(* IEC 61131-3 sources: daoli-st-library/DL_Device (part 18) *)

(* ---- FB_DL_CrystallizerVacuumCtrl.st ---- *)
(*
  Component : FB_DL_CrystallizerVacuumCtrl
  Category  : DL_Device
  Type      : FB
  Complexity: C2
  VERSION   : v1.0.0
  功能      : 结晶罐真空控制：ENUM 四态（Off/Run/Lost/Fault），真空泵按压差分级投运，按锤度算沸点升高与罐内沸点，真空丢失延时联锁停泵。
  开源溯源  : 道莅原创 clean-room 自研（无外部代码引用）｜License: MIT
  边界条件  : ① 真空度输入按罐内绝对压力定义 [kPa]：实测值升高即真空丢失，判据方向不得反接；
              ② 沸点升高按 锤度/(100-锤度) 经验式，锤度须 < 100 °Bx 且钳位 0~30 K；
              ③ 真空丢失锁存后全泵切除（防倒吸油返），唯一解除路径 = bReset 上升沿。
*)

TYPE E_DL_VacMode :
(
    eOff   := 0,    (* 停机：使能撤销 / Off, disabled *)
    eRun   := 10,   (* 运行：分级投运 / Running with staged pumps *)
    eLost  := 20,   (* 真空丢失：全泵切除锁存 / Vacuum lost, pumps cut off *)
    eFault := 90    (* 故障：锁存待复位 / Fault latched *)
);
END_TYPE

FUNCTION_BLOCK FB_DL_CrystallizerVacuumCtrl
VAR_INPUT
    bEnable     : BOOL;   (* 使能电平 [-] Enable level *)
    bReset      : BOOL;   (* 复位上升沿，清丢失与故障锁存 [-] Reset edge *)
    fVacuumKPa  : REAL;   (* 罐内绝对压力实测 [kPa] Measured absolute pressure *)
    fVacSetKPa  : REAL;   (* 目标绝对压力设定 [kPa] Absolute pressure setpoint *)
    fVacLostKPa : REAL;   (* 真空丢失判据压力 [kPa] Vacuum-lost pressure threshold *)
    fBrixPct    : REAL;   (* 糖膏锤度 [°Bx] Massecuite brix *)
    fWaterBoilC : REAL;   (* 当前真空下纯水沸点 [°C] Water boiling point at this vacuum *)
    tLostDelay  : TIME;   (* 真空丢失确认延时 [ms] Vacuum-lost confirmation delay *)
    nPumpMax    : INT;    (* 可用真空泵台数 1~3 [-] Available pump count *)
END_VAR
VAR_OUTPUT
    abPumpCmd  : ARRAY[0..2] OF BOOL;  (* 三级真空泵指令 [-] Vacuum pump commands *)
    nPumpRun   : INT;                  (* 当前投运泵台数 [-] Running pump count *)
    fBoilRiseK : REAL;                 (* 沸点升高 [K] Boiling point elevation *)
    fBoilTempC : REAL;                 (* 罐内糖膏沸点 [°C] Massecuite boiling point *)
    bVacLost   : BOOL;                 (* 真空丢失锁存标志 [-] Vacuum lost latch *)
    eMode      : E_DL_VacMode;         (* 模式出口，段尾单点映射 [-] Mode outlet *)
    bError     : BOOL;                 (* 故障锁存标志 [-] Fault latch flag *)
    uErrId     : UDINT;                (* 事件码，0 = 无事件 [-] Event code *)
END_VAR
VAR
    rtReset  : R_TRIG;   (* 复位沿实例，每拍无条件刷新 / Reset edge *)
    tonLost  : TON;      (* 真空丢失确认计时 / Vacuum lost timer *)
    _eMode   : E_DL_VacMode := E_DL_VacMode.eOff;  (* 内部模式 / Internal mode *)
    _bLost   : BOOL;     (* 真空丢失锁存位（锁存量） / Latched vacuum lost bit *)
    _bFault  : BOOL;     (* 故障锁存位（锁存量） / Latched fault bit *)
    _uFault  : UDINT;    (* 故障码锁存（锁存量） / Latched fault code *)
    _bCfgBad : BOOL;     (* 组态非法当拍量 [-] Config illegal flag *)
    _bNonFin : BOOL;     (* 输入非有限当拍量 [-] Non-finite input flag *)
    nIdx     : INT;      (* 泵组遍历下标 [-] Pump loop index *)
    fErrKPa  : REAL;     (* 压差（实测 - 设定） [kPa] Pressure error *)
    fDenBrix : REAL;     (* 锤度余量（100 - 锤度） [°Bx] Brix headroom *)
END_VAR
VAR CONSTANT
    DL_EPS      : REAL := 1.0E-9;   (* 除零判定容差 [无量纲] Divide-by-zero tolerance *)
    DL_BAND1    : REAL := 1.0;      (* 一级投运压差 [kPa] Stage 1 pressure band *)
    DL_BAND2    : REAL := 4.0;      (* 二级投运压差 [kPa] Stage 2 pressure band *)
    DL_BAND3    : REAL := 8.0;      (* 三级投运压差 [kPa] Stage 3 pressure band *)
    DL_RISE_K   : REAL := 2.6;      (* 沸点升高经验系数 [K] Elevation coefficient *)
    DL_RISE_MAX : REAL := 30.0;     (* 沸点升高上限 [K] Elevation upper clamp *)
    DL_PCT_BASE : REAL := 100.0;    (* 百分比基准 [°Bx 基准] Percent base *)
    DL_IDX_MAX  : INT := 2;         (* 泵组最高下标 [-] Highest pump index *)
END_VAR

(* —— 段 0｜沿与定时器每拍无条件刷新（禁置于 IF/CASE 内，使能挂 IN 引脚） —— *)
rtReset(CLK := bReset);
tonLost(IN := bEnable AND (fVacuumKPa >= fVacLostKPa) AND (NOT _bLost), PT := tLostDelay);

(* —— 段 1｜每拍量预清零 + 泵指令全预置（锁存量 _bLost/_bFault/_uFault 不入清单） —— *)
uErrId := 16#0000_0000;
_bCfgBad := FALSE;
_bNonFin := FALSE;
nPumpRun := 0;
FOR nIdx := 0 TO 2 DO
    IF (nIdx >= 0) AND (nIdx <= DL_IDX_MAX) THEN
        abPumpCmd[nIdx] := FALSE;            (* 泵指令预置停止 [-] / Pump preset off *)
    END_IF
END_FOR

(* —— 段 2｜非有限拦截与组态闸（覆盖压力设定/丢失判据/锤度/延时/泵数） —— *)
IF (fVacuumKPa <> fVacuumKPa) OR ((fVacuumKPa - fVacuumKPa) <> 0.0)
   OR (fBrixPct <> fBrixPct) OR ((fBrixPct - fBrixPct) <> 0.0)
   OR (fVacSetKPa <> fVacSetKPa) OR ((fVacSetKPa - fVacSetKPa) <> 0.0)
   OR (fVacLostKPa <> fVacLostKPa) OR ((fVacLostKPa - fVacLostKPa) <> 0.0)
   OR (fWaterBoilC <> fWaterBoilC) OR ((fWaterBoilC - fWaterBoilC) <> 0.0) THEN
    _bNonFin := TRUE;
END_IF
IF (fVacSetKPa <= DL_EPS) OR (fVacLostKPa <= fVacSetKPa) OR (tLostDelay = T#0S)
   OR (nPumpMax < 1) OR (nPumpMax > 3) OR (fBrixPct < 0.0) OR (fBrixPct >= DL_PCT_BASE) THEN
    _bCfgBad := TRUE;
END_IF

(* —— 段 3｜沸点升高与罐内沸点：dT = 2.6·B/(100-B)，钳位 0~30 K —— *)
fDenBrix := DL_PCT_BASE - fBrixPct;
IF fDenBrix > DL_EPS THEN
    fBoilRiseK := DL_RISE_K * fBrixPct / fDenBrix;
ELSE
    fBoilRiseK := DL_RISE_MAX;               (* 锤度近饱和：按上限处理 *)
END_IF
IF fBoilRiseK < 0.0 THEN
    fBoilRiseK := 0.0;
ELSIF fBoilRiseK > DL_RISE_MAX THEN
    fBoilRiseK := DL_RISE_MAX;
END_IF
fBoilTempC := fWaterBoilC + fBoilRiseK;

(* —— 段 4｜复位沿：一次性清丢失与故障锁存（唯一解除路径，恒可达） —— *)
IF rtReset.Q THEN
    _bLost := FALSE;
    _bFault := FALSE;
    _uFault := 16#0000_0000;
    _eMode := E_DL_VacMode.eOff;
END_IF
IF _bCfgBad AND (NOT _bFault) THEN
    _bFault := TRUE;
    _uFault := 16#0029_0001;                 (* 故障级：组态非法 / Fault code bad config *)
END_IF
IF _bNonFin AND (NOT _bFault) THEN
    _bFault := TRUE;
    _uFault := 16#0029_0002;                 (* 故障级：压力或锤度非有限 / Non-finite input *)
END_IF
IF tonLost.Q AND (NOT _bLost) THEN
    _bLost := TRUE;                          (* 真空丢失锁存：全泵切除防倒吸 *)
END_IF

(* —— 段 5｜模式机：四态全覆盖 + ELSE 兜底 —— *)
CASE _eMode OF
E_DL_VacMode.eOff:
    nPumpRun := 0;
    IF bEnable AND (NOT _bLost) AND (NOT _bFault) AND (NOT _bCfgBad) AND (NOT _bNonFin) THEN
        _eMode := E_DL_VacMode.eRun;         (* 迁入条件：使能且无任何锁存 *)
    END_IF

E_DL_VacMode.eRun:
    (* 压差分级投运：实测绝对压力高于设定越多，投运泵台数越多 *)
    fErrKPa := fVacuumKPa - fVacSetKPa;
    IF fErrKPa > DL_BAND3 THEN
        nPumpRun := 3;
    ELSIF fErrKPa > DL_BAND2 THEN
        nPumpRun := 2;
    ELSIF fErrKPa > DL_BAND1 THEN
        nPumpRun := 1;
    ELSE
        nPumpRun := 0;
    END_IF
    IF nPumpRun > nPumpMax THEN
        nPumpRun := nPumpMax;                (* 受可用台数限制 [-] / Limited by available pumps *)
    END_IF
    IF _bLost THEN
        _eMode := E_DL_VacMode.eLost;        (* 迁出条件 1：真空丢失 *)
    ELSIF _bFault THEN
        _eMode := E_DL_VacMode.eFault;       (* 迁出条件 2：故障锁存 *)
    ELSIF NOT bEnable THEN
        _eMode := E_DL_VacMode.eOff;         (* 迁出条件 3：使能撤销 *)
    END_IF

E_DL_VacMode.eLost:
    nPumpRun := 0;                           (* 丢失相：全泵切除（防倒吸油返） *)
    IF NOT _bLost THEN
        _eMode := E_DL_VacMode.eOff;         (* 迁出条件：锁存被复位沿清除 *)
    END_IF

E_DL_VacMode.eFault:
    nPumpRun := 0;                           (* 故障相：全泵切除 *)
    IF (NOT _bFault) AND (NOT _bLost) THEN
        _eMode := E_DL_VacMode.eOff;         (* 迁出条件：故障锁存被复位沿清除 *)
    END_IF

ELSE
    _bFault := TRUE;                         (* 兜底：非法模式锁存 *)
    _uFault := 16#0029_0009;
    _eMode := E_DL_VacMode.eFault;
END_CASE

(* —— 段 6｜泵指令下发：仅运行相按台数投运，其余相全切除 —— *)
IF _eMode = E_DL_VacMode.eRun THEN
    FOR nIdx := 0 TO 2 DO
        IF (nIdx >= 0) AND (nIdx <= DL_IDX_MAX) THEN
            abPumpCmd[nIdx] := nIdx < nPumpRun;   (* 前 nPumpRun 台投运 [-] / First N pumps on *)
        END_IF
    END_FOR
ELSE
    nPumpRun := 0;
END_IF

(* —— 段 7｜出口单点映射 —— *)
eMode := _eMode;
bVacLost := _bLost;
bError := _bFault;
IF _bFault AND (_uFault <> 16#0000_0000) THEN
    uErrId := _uFault;                       (* 故障码锁存回放 / Latched fault replay *)
END_IF
END_FUNCTION_BLOCK

(* ---- FB_DL_CurtainEFEMZone.st ---- *)
(*
  FB_DL_CurtainEFEMZone  —  EFEM 区内光幕分区（四路遮光判向 / 屏蔽窗管理 / 顺序故障锁存）/ EFEM zone light-curtain muting
  分类 Category : DL_Device
  码位 Code     : 16#03_2_0C
  版本 Version  : 1.0.2
  来源 Source   : t1-5-tcopen — IEC 61131-3 标准语义的道莅防御性实现
  溯源 Origin   : TwinCAT/TCopen 光幕屏蔽（muting）公开语义借鉴，clean-room 实现，未复制任何源码行
  功能 Function : 1) 四路光幕（进入侧 A / 进入侧 B / 区内 C / 出口侧 D）逐拍采集 bClear / bFault；
                  2) 遮光事件（上升沿）按先后入序列缓冲，A→B→C→D 判「正向通过」，D→C→B→A 判「反向通过」；
                  3) 序列至少两路且方向已定才允许开屏蔽窗（bMutingActive），屏蔽窗受 tMutingMax 强制限时；
                  4) 屏蔽期与非屏蔽期**都**输出受控速度限幅 fSpeedLimitOut（屏蔽 ≠ 无限速，规格强制项）；
                  5) 非顺序遮光（如 C 先于 A）或相邻遮光间隔超 tSequenceGap → bSequenceFault 锁存并禁屏蔽。
  边界 Boundary : ① 任一传感器自检失败（bFault = TRUE）**立即退出屏蔽**并置 023C（不得静默屏蔽，安全侧）；
                  ② tMutingMax 到点强制解屏蔽并置 022C（屏蔽超时是故障级，必须人工确认后复位）；
                  ③ 判向超 tSequenceGap 判「顺序失败」而非「无事件」：间隔超限说明通过节奏异常（可能是爬行/滞留），
                     按失败处理并清序列缓冲，码 012C（信息级）+ 021C（故障级，仅非顺序时）；
                     间隙计时随每次新遮光事件重启，间隔判据对每一对相邻事件均生效（R38 返修口径）；
                  ④ 解除式自证：bSequenceFault 解除 = bReset AND NOT bMutingEnable（组态退出屏蔽即可满足，R28-1）；
                     022C / 023C 同样由 rtReset.Q 清除，与本条互不掩盖（R188 双路径）；
                  ⑤ bZoneSafe 语义：区内光幕 C 通光，或屏蔽窗合法开启且无顺序故障与无传感器自检失败；
                     其余一律 FALSE（含 eAborted / eFault 相），上层据此做区域降速或停车；
                  ⑥ 时间参数 <= 0、速度限幅 <= 0、tSequenceGap > tMutingMax 均判组态错 020C（后者会让
                     屏蔽窗在序列判向前就超时，属不可能组态）。
  依赖 Depends  : I_DL_LightCurtain（DL_Device 既有契约，×4 注入，不实例化）；
                  仅 Standard.library（TON / R_TRIG / ABS / MIN / MAX）
  同拍双窗配比  : tSequenceGap（相邻遮光间隔）与 tMutingMax（屏蔽窗总时长）同源于通过节奏；
                  配比约束 tSequenceGap <= tMutingMax（组态闸强制），保证序列判据不会晚于屏蔽窗失效

  码表 Error codes（本件格 03_2_0C，子码步进 +0x10）:
    16#0003_020C 故障级：组态非法（时间参数 <= 0 / 速度限幅 <= 0 / tSequenceGap > tMutingMax）
    16#0003_021C 故障级：遮光顺序故障（非顺序遮光，锁存并禁屏蔽）
    16#0003_022C 故障级：屏蔽超时（tMutingMax 到点强制解屏蔽，锁存）
    16#0003_023C 故障级：光幕传感器自检失败（立即退出屏蔽，锁存）
    16#0003_024C 故障级：状态机落 ELSE 兜底（非法相位 ID）
    16#0003_010C 信息级：屏蔽窗开启（序列成立且方向已定，不置 bError）
    16#0003_011C 信息级：屏蔽窗正常结束（序列走完或全部通光，不置 bError）
    16#0003_012C 信息级：相邻遮光间隔超 tSequenceGap，序列缓冲已清（判向失败，不置 bError）

  修订历史 Revision :
    2026-11-18  v1.0.0  R37 首版
    2026-11-18  v1.0.2  R38 返修：间隙计时随新遮光事件重启（_bGapBreak 断输入请求，R188 自复位范式），间隔判据对每一对相邻事件均生效
  R38 已修复    : R37 终审挂账「间隙计时器不随新遮光事件重启」已修复（四路遮光上升沿统一汇合点置 _bGapBreak）
*)

TYPE E_DL_MutingState :
(
    eIdle     := 0,   // 空闲：未使能或屏蔽功能关闭 / Idle, muting disabled by the master enable or the configuration
    eEval     := 10,  // 评估：等待首个遮光事件 / Evaluating, waiting for the first occlusion
    eSeqCheck := 20,  // 判向：已有一路遮光，等第二路定方向 / Sequence check, waiting for the second occlusion
    eMuting   := 30,  // 屏蔽中：屏蔽窗开启并限时 / Muting, the window is open and time-limited
    eAborted  := 40,  // 中止：屏蔽被超时/自检失败中止，等待复位 / Aborted, waiting for a reset
    eFault    := 90   // 故障：顺序故障或组态故障锁定 / Fault, a latched sequence or configuration fault
);
END_TYPE

FUNCTION_BLOCK FB_DL_CurtainEFEMZone
VAR_INPUT
    bEnable       : BOOL := FALSE;             // 总使能，FALSE 时禁屏蔽并回空闲 / Master enable, low level forbids muting
    bReset        : BOOL := FALSE;             // 复位，上升沿清故障锁存 / Reset, rising edge clears the latch
    bMutingEnable : BOOL := FALSE;             // 屏蔽功能组态使能（退出即解除顺序故障）/ Muting feature enable
    fZoneSpeedLimit : REAL := 300.0;           // 区内速度限幅 [mm/s]，域 > 0 / Zone speed limit [mm/s]
    tMutingMax    : TIME := T#30S;             // 屏蔽最长时限 [ms]，域 > 0 / Maximum muting duration [ms]
    tSequenceGap  : TIME := T#5S;              // 相邻遮光间隔上限 [ms]，域 > 0 且 <= tMutingMax / Adjacent occlusion gap [ms]
    tClearHold    : TIME := T#500MS;           // 全通光确认驻留 [ms]，域 > 0 / All-clear confirm dwell [ms]
END_VAR
VAR_OUTPUT
    bZoneSafe      : BOOL;                     // 区域安全（区内无人或屏蔽合法）/ Zone safe
    bMutingActive  : BOOL;                     // 屏蔽进行中 / Muting active
    bSequenceFault : BOOL;                     // 遮光顺序故障锁存 / Occlusion sequence fault latched
    bMutingTimeout : BOOL;                     // 屏蔽超时锁存 / Muting timeout latched
    bSensorFault   : BOOL;                     // 任一光幕自检失败 / Any curtain self-test failure
    fSpeedLimitOut : REAL;                     // 生效速度限幅 [mm/s]（屏蔽期同样受控）/ Effective speed limit [mm/s]
    nSeqLength     : INT;                      // 当前序列长度 [路] / Present sequence length
    bValid         : BOOL;                     // 判据可用标志 / Criteria usable
    bError         : BOOL;                     // 故障标志，派生自锁存 / Fault flag derived from the latch
    nErrId         : UDINT;                    // 事件码，0 = 无事件 / Event code, 0 = no event
    eStateOut      : E_DL_MutingState;         // 状态出口，段尾单点映射 / State outlet, mapped at the tail
END_VAR
VAR_IN_OUT
    iCurtainA : I_DL_LightCurtain;             // 进入侧 A 光幕引用（注入，不实例化）/ Entry side A curtain reference
    iCurtainB : I_DL_LightCurtain;             // 进入侧 B 光幕引用（注入，不实例化）/ Entry side B curtain reference
    iCurtainC : I_DL_LightCurtain;             // 区内 C 光幕引用（注入，不实例化）/ In-zone C curtain reference
    iCurtainD : I_DL_LightCurtain;             // 出口侧 D 光幕引用（注入，不实例化）/ Exit side D curtain reference
END_VAR
VAR
    tonMuting   : TON;                         // 屏蔽最长时限计时，每拍无条件调用 / Muting duration timer, called unconditionally
    tonGap      : TON;                         // 相邻遮光间隔计时，每拍无条件调用 / Occlusion gap timer, called unconditionally
    tonClear    : TON;                         // 全通光确认驻留，每拍无条件调用 / All-clear dwell timer, called unconditionally
    tonHeart    : TON;                         // 周期心跳窗，自复位 / Periodic heartbeat window, self-resetting
    rtReset     : R_TRIG;                      // 复位上升沿 / Reset rising edge
    rtA         : R_TRIG;                      // A 路遮光上升沿 / Curtain A occlusion edge
    rtB         : R_TRIG;                      // B 路遮光上升沿 / Curtain B occlusion edge
    rtC         : R_TRIG;                      // C 路遮光上升沿 / Curtain C occlusion edge
    rtD         : R_TRIG;                      // D 路遮光上升沿 / Curtain D occlusion edge
    _eState     : E_DL_MutingState := E_DL_MutingState.eIdle;  // 内部相位（CASE 唯一写入目标）/ Internal phase
    _uFault     : UDINT;                       // 故障码锁存 / Latched fault code
    _uInfo      : UDINT;                       // 信息码，每拍重算 / Information code, recomputed per scan
    _bFault     : BOOL;                        // 故障锁存位 / Latched fault bit
    _bCfgBad    : BOOL;                        // 组态非法聚合 / Configuration invalid aggregate
    _bOccA      : BOOL;                        // A 路遮光 / Curtain A occluded
    _bOccB      : BOOL;                        // B 路遮光 / Curtain B occluded
    _bOccC      : BOOL;                        // C 路遮光 / Curtain C occluded
    _bOccD      : BOOL;                        // D 路遮光 / Curtain D occluded
    _bAnyOcc    : BOOL;                        // 任一路遮光 / Any curtain occluded
    _bAllClear  : BOOL;                        // 全部通光 / All curtains clear
    _bSensFault : BOOL;                        // 传感器自检失败聚合 / Sensor self-test failure aggregate
    _bSeqFault  : BOOL;                        // 顺序故障保持量 / Held sequence fault
    _bTimeout   : BOOL;                        // 屏蔽超时保持量 / Held muting timeout
    _bNewEvent  : BOOL;                        // 本拍有新的遮光事件 / A new occlusion event occurred
    _bGapBroken : BOOL;                        // 相邻间隔超限 / The gap limit was violated
    _bGapBreak  : BOOL := FALSE;               // 间隙计时断输入请求（新遮光事件沿触发，R188 自复位范式）/ Gap-timer break request, set by a new occlusion edge
    _nNewIdx    : INT;                         // 本拍新事件的序号（A=1..D=4）/ Order index of the new event
    _nDir       : INT;                         // 判向结果（0 未知 / +1 正向 / −1 反向）/ Direction verdict
    _anSeq      : ARRAY[0..3] OF INT;          // 序列缓冲（存序号 1..4）[路] / Sequence buffer holding indices one to four
    _nSeqLen    : INT;                         // 序列长度 [路] / Sequence length
    _nLastIdx   : INT;                         // 序列末项序号 / Index of the last accepted event
    _bHeartBrk  : BOOL := TRUE;                // 心跳窗断输入一拍 / One-scan heartbeat break
END_VAR
VAR CONSTANT
    DL_IDX_A      : INT := 1;          // A 路序号（进入侧）/ Order index of curtain A
    DL_IDX_B      : INT := 2;          // B 路序号（进入侧）/ Order index of curtain B
    DL_IDX_C      : INT := 3;          // C 路序号（区内）/ Order index of curtain C
    DL_IDX_D      : INT := 4;          // D 路序号（出口侧）/ Order index of curtain D
    DL_SEQ_NONE   : INT := 0;          // 序列空 / Empty sequence marker
    DL_SPEED_MIN  : REAL := 1.0;       // 速度限幅下限 [mm/s]（0 会让轴失去使能语义）/ Speed limit floor
    DL_SPEED_MAX  : REAL := 5000.0;    // 速度限幅上限 [mm/s] / Speed limit ceiling
    DL_HEART_WINDOW : TIME := T#2S;    // 心跳观察窗 [ms]，自复位节拍 / Heartbeat window, self-resetting
END_VAR

(* —— 段 0：定时器与边缘检测无条件周期刷新（R182：调用语句不得置于 IF / CASE 内） —— *)
rtReset(CLK := bReset);                                          // 复位上升沿，每拍必调
rtA(CLK := _bOccA);                                              // A 路遮光上升沿，每拍必调
rtB(CLK := _bOccB);                                              // B 路遮光上升沿，每拍必调
rtC(CLK := _bOccC);                                              // C 路遮光上升沿，每拍必调
rtD(CLK := _bOccD);                                              // D 路遮光上升沿，每拍必调
tonHeart(IN := (NOT tonHeart.Q) AND (NOT _bHeartBrk), PT := DL_HEART_WINDOW);  // 心跳窗自复位
_bHeartBrk := FALSE;                                             // 断输入拍在调用后自清
tonMuting(IN := (_eState = E_DL_MutingState.eMuting), PT := tMutingMax);        // 屏蔽限时（表达式入参）
tonGap(IN := ((_nSeqLen > 0) AND (_nSeqLen < 4)) AND (NOT _bGapBreak), PT := tSequenceGap);  // 相邻遮光间隔（表达式入参；断输入请求使 ET 随新事件归零重启）
_bGapBreak := FALSE;                                             // 断输入拍在调用后自清（新遮光沿在段 5 置位）
tonClear(IN := _bAllClear, PT := tClearHold);                                   // 全通光确认驻留（表达式入参）

(* —— 段 1：单拍量预清零（序列缓冲 / 保持量 / 锁存不入清单，R187①） —— *)
_uInfo      := 16#0000_0000;   // 信息码每拍重算
bError      := FALSE;          // 故障出口每拍重算，段 8 由锁存派生
bValid      := FALSE;          // 可用标志缺省 FALSE
bMutingActive := FALSE;        // 屏蔽出口缺省 FALSE，段 8 单点置位
bZoneSafe   := FALSE;          // 区域安全缺省 FALSE（安全侧缺省）
_bCfgBad    := FALSE;          // 组态非法预清零
_bNewEvent  := FALSE;          // 新事件标志预清零
_bGapBroken := FALSE;          // 间隔超限标志预清零
_nNewIdx    := DL_SEQ_NONE;    // 新事件序号预清零

(* —— 段 2：复位沿清锁存 + 按码专清（R188 双路径，互不掩盖） —— *)
IF rtReset.Q THEN
    IF NOT bMutingEnable THEN
        _bSeqFault := FALSE;           // 解除式：bReset AND NOT bMutingEnable（组态退出屏蔽即可满足）
    END_IF
    IF NOT _bSeqFault THEN
        _bFault   := FALSE;            // 顺序故障保持量已释放才清故障位（防「码清位不清」）
        _uFault   := 16#0000_0000;     // 清锁存码
        _bTimeout := FALSE;            // 屏蔽超时保持量清零（与 022C 同源）
        _nSeqLen  := 0;                // 序列缓冲长度归零
        _nDir     := 0;                // 判向结果归零
    END_IF
END_IF
IF (_uFault = 16#0003_021C) AND (NOT _bSeqFault) THEN
    _uFault := 16#0000_0000;           // 按码专清：顺序故障保持量已释放 → 对应码清除
    _bFault := FALSE;                  // 锁存位同步清
END_IF
IF (_uFault = 16#0003_022C) AND (NOT _bTimeout) THEN
    _uFault := 16#0000_0000;           // 按码专清：屏蔽超时保持量已释放 → 对应码清除
    _bFault := FALSE;                  // 锁存位同步清
END_IF

(* —— 段 3：组态域闸（覆盖全部参与判据换算的引脚，R151） —— *)
IF (fZoneSpeedLimit <> fZoneSpeedLimit) OR (fZoneSpeedLimit < DL_SPEED_MIN) THEN
    _bCfgBad := TRUE;              // 速度限幅非法（下限防 0 值让上层误判为无限速）
END_IF
IF fZoneSpeedLimit > DL_SPEED_MAX THEN
    _bCfgBad := TRUE;              // 速度限幅超上界（组态量纲错）
END_IF
IF TIME_TO_DINT(tMutingMax) <= 0 THEN
    _bCfgBad := TRUE;              // 屏蔽限时非法
END_IF
IF TIME_TO_DINT(tSequenceGap) <= 0 THEN
    _bCfgBad := TRUE;              // 判向间隔非法
END_IF
IF TIME_TO_DINT(tClearHold) <= 0 THEN
    _bCfgBad := TRUE;              // 全通光确认驻留非法
END_IF
IF (TIME_TO_DINT(tSequenceGap) > 0) AND (TIME_TO_DINT(tMutingMax) > 0) AND
   (TIME_TO_DINT(tSequenceGap) > TIME_TO_DINT(tMutingMax)) THEN
    _bCfgBad := TRUE;              // 判向间隔大于屏蔽限时：序列判据必然晚于屏蔽窗失效（不可能组态）
END_IF
IF _bCfgBad THEN
    _uFault := 16#0003_020C;       // 故障级：组态非法
    _bFault := TRUE;               // 锁存位置位（复位沿可清）
    bError  := TRUE;               // 故障标志置位（R45 配对）
    _eState := E_DL_MutingState.eFault;  // 进故障相
END_IF

(* —— 段 4：四路光幕采集（只读属性，零命令下发） —— *)
_bOccA := NOT iCurtainA.bClear;    // A 路遮光（通光取反）
_bOccB := NOT iCurtainB.bClear;    // B 路遮光
_bOccC := NOT iCurtainC.bClear;    // C 路遮光（区内）
_bOccD := NOT iCurtainD.bClear;    // D 路遮光
_bAnyOcc := _bOccA OR _bOccB OR _bOccC OR _bOccD;                    // 任一路遮光
_bAllClear := (NOT _bAnyOcc);                                       // 全部通光
_bSensFault := iCurtainA.bFault OR iCurtainB.bFault OR
               iCurtainC.bFault OR iCurtainD.bFault;                // 任一路自检失败
bSensorFault := _bSensFault;                                        // 自检失败出口（安全镜像）

(* —— 段 4A：自检失败立即退出屏蔽（安全侧，先于一切序列判定，R190 归因唯一） —— *)
IF _bSensFault THEN
    IF (_eState = E_DL_MutingState.eMuting) OR (_eState = E_DL_MutingState.eSeqCheck) THEN
        _uFault := 16#0003_023C;   // 故障级：光幕传感器自检失败，屏蔽立即退出
        _bFault := TRUE;           // 锁存
        bError  := TRUE;           // 故障标志置位（R45 配对）
        _eState := E_DL_MutingState.eAborted;  // 中止相（等复位）
        _nSeqLen := 0;             // 序列缓冲清空（自检失败后旧序列不可信）
        _nDir := 0;                // 判向清空
    END_IF
END_IF

(* —— 段 5：遮光事件排序（序号入缓冲，方向唯一确定后才允许屏蔽） —— *)
IF _bAnyOcc AND (NOT _bSensFault) THEN
    IF rtA.Q THEN
        _bNewEvent := TRUE; _nNewIdx := DL_IDX_A;   // A 路新事件
    ELSIF rtB.Q THEN
        _bNewEvent := TRUE; _nNewIdx := DL_IDX_B;   // B 路新事件
    ELSIF rtC.Q THEN
        _bNewEvent := TRUE; _nNewIdx := DL_IDX_C;   // C 路新事件
    ELSIF rtD.Q THEN
        _bNewEvent := TRUE; _nNewIdx := DL_IDX_D;   // D 路新事件
    END_IF
END_IF

IF _bNewEvent THEN
    _bGapBreak := TRUE;                             // R38 返修：新遮光上升沿（A/B/C/D 四路统一汇合点）置断输入请求，
                                                    // 下一拍 tonGap IN 断开（Q 天然为 FALSE）→ ET 归零，间隙从新事件重新计时；
                                                    // 本拍 _bGapBreak 置位不影响本拍已完成的 tonGap 调用（段 0 先行）
    IF tonGap.Q AND (_nSeqLen > 0) THEN
        _bGapBroken := TRUE;                        // 相邻遮光间隔超限：判向失败（不是「无事件」）
        _nSeqLen := 0;                              // 序列缓冲清空
        _nDir := 0;                                 // 方向作废
        _uInfo := 16#0003_012C;                     // 信息级：间隔超限，序列已清
    END_IF
    IF _nSeqLen = 0 THEN
        _anSeq[0] := _nNewIdx;                      // 首路遮光入缓冲
        _nSeqLen := 1;                              // 长度 1
        _nLastIdx := _nNewIdx;                      // 末项记录
        _nDir := 0;                                 // 方向待定
    ELSIF _nSeqLen < 4 THEN
        IF _nDir = 0 THEN
            IF _nNewIdx = (_nLastIdx + 1) THEN
                _nDir := 1;                         // 序号递增：正向通过
            ELSIF _nNewIdx = (_nLastIdx - 1) THEN
                _nDir := -1;                        // 序号递减：反向通过
            ELSE
                _bSeqFault := TRUE;                 // 非相邻：非顺序遮光（如 C 先于 A）
            END_IF
        ELSE
            IF _nNewIdx <> (_nLastIdx + _nDir) THEN
                _bSeqFault := TRUE;                 // 与已定方向不符：非顺序遮光
            END_IF
        END_IF
        IF _bSeqFault THEN
            _uFault := 16#0003_021C;                // 故障级：遮光顺序故障（禁屏蔽）
            _bFault := TRUE;                        // 锁存
            bError  := TRUE;                        // 故障标志置位（R45 配对）
            _eState := E_DL_MutingState.eFault;     // 进故障相
        ELSE
            _anSeq[_nSeqLen] := _nNewIdx;           // 顺序成立：事件入缓冲
            _nSeqLen := _nSeqLen + 1;               // 长度递增（上限 4 由外条件守）
            _nLastIdx := _nNewIdx;                  // 末项更新
        END_IF
    END_IF
END_IF
nSeqLength := _nSeqLen;                             // 序列长度出口（诊断用）

(* —— 段 6：相位机（只做迁移；屏蔽出口在段 8） —— *)
CASE _eState OF

E_DL_MutingState.eIdle:
    IF bEnable AND bMutingEnable AND (NOT _bFault) AND (NOT _bCfgBad) THEN
        _eState := E_DL_MutingState.eEval;          // 使能且屏蔽功能开：进评估相
    END_IF

E_DL_MutingState.eEval:
    IF (NOT bEnable) OR (NOT bMutingEnable) THEN
        _eState := E_DL_MutingState.eIdle;          // 退出屏蔽功能：回空闲
    ELSIF _nSeqLen >= 1 THEN
        _eState := E_DL_MutingState.eSeqCheck;      // 已有首路遮光：进判向相
    END_IF

E_DL_MutingState.eSeqCheck:
    IF (NOT bEnable) OR (NOT bMutingEnable) THEN
        _eState := E_DL_MutingState.eIdle;          // 退出屏蔽功能
        _nSeqLen := 0;                              // 序列清空
        _nDir := 0;                                 // 方向清空
    ELSIF (_nSeqLen >= 2) AND (_nDir <> 0) THEN
        _eState := E_DL_MutingState.eMuting;        // 方向已定：开屏蔽窗
        _uInfo  := 16#0003_010C;                    // 信息级：屏蔽窗开启
    ELSIF tonGap.Q THEN
        _uInfo := 16#0003_012C;                     // 信息级：判向超时（不足两路）
        _nSeqLen := 0;                              // 序列清空，等下一轮
        _nDir := 0;
        _eState := E_DL_MutingState.eEval;          // 回评估相
    END_IF

E_DL_MutingState.eMuting:
    IF _bSensFault THEN
        _eState := E_DL_MutingState.eAborted;       // 自检失败：立即退出（段 4A 已置码）
    ELSIF (NOT bEnable) OR (NOT bMutingEnable) THEN
        _eState := E_DL_MutingState.eEval;          // 组态退出屏蔽：解屏蔽
        _nSeqLen := 0;
        _nDir := 0;
    ELSIF tonMuting.Q THEN
        _bTimeout := TRUE;                          // 屏蔽超时保持量
        _uFault := 16#0003_022C;                    // 故障级：屏蔽超时强制解屏蔽
        _bFault := TRUE;                            // 锁存
        bError  := TRUE;                            // 故障标志置位（R45 配对）
        _eState := E_DL_MutingState.eAborted;       // 中止相
        _nSeqLen := 0;
        _nDir := 0;
    ELSIF tonClear.Q THEN
        _uInfo := 16#0003_011C;                     // 信息级：全部通光并驻留完成，屏蔽窗正常结束
        _nSeqLen := 0;                              // 序列清空，准备下一件
        _nDir := 0;
        _eState := E_DL_MutingState.eEval;          // 回评估相
    END_IF

E_DL_MutingState.eAborted:
    IF (NOT bEnable) THEN
        _eState := E_DL_MutingState.eIdle;          // 失能：回空闲
    ELSIF (NOT _bFault) AND bMutingEnable AND (NOT _bSensFault) THEN
        _eState := E_DL_MutingState.eEval;          // 复位完成且自检恢复：回评估相
    END_IF

E_DL_MutingState.eFault:
    IF (NOT _bFault) AND (NOT _bCfgBad) AND bEnable AND bMutingEnable THEN
        _eState := E_DL_MutingState.eEval;          // 锁存已清且组态合法：回评估相
    END_IF

ELSE
    _uFault := 16#0003_024C;                        // 故障级：相位 ID 越界（枚举兜底）
    _bFault := TRUE;                                // 锁存
    bError  := TRUE;                                // 故障标志置位（R45 配对）
    _eState := E_DL_MutingState.eFault;             // 强制回故障相
END_CASE

(* —— 段 7：故障码优先级链（每个 bError 置位源在此均有码，R45 配对） —— *)
IF _bCfgBad THEN
    bError := TRUE;                                 // 组态非法：码已在段 3 置位（020C）
END_IF

(* —— 段 8：出口单点映射（名实同源；锁存码回放，禁同拍抹除） —— *)
bMutingActive   := (_eState = E_DL_MutingState.eMuting) AND (NOT _bFault);  // 屏蔽出口：仅在屏蔽相且无故障
bSequenceFault  := _bSeqFault;                                              // 顺序故障出口（保持量）
bMutingTimeout  := _bTimeout;                                               // 屏蔽超时出口（保持量）
fSpeedLimitOut  := fZoneSpeedLimit;                                         // 生效限幅：屏蔽期同样受控（屏蔽 ≠ 无限速）
bZoneSafe       := ((NOT _bOccC) AND (NOT _bSensFault) AND (NOT _bFault)) OR
                   (bMutingActive AND (NOT _bSeqFault) AND (NOT _bSensFault));  // 区域安全：区内通光或屏蔽合法
eStateOut       := _eState;                                                 // 状态出口
IF _bFault THEN
    nErrId := _uFault;                           // 故障锁存码回放（不在故障相按当下输入重推）
    bError := TRUE;                              // 故障出口派生自锁存
ELSE
    nErrId := _uInfo;                            // 信息码
END_IF
bValid := bEnable AND bMutingEnable AND (NOT _bFault) AND (NOT _bCfgBad);  // 判据可用

END_FUNCTION_BLOCK

(* ---- FB_DL_CylStrokeTimeBank.st ---- *)
(*==============================================================================
 * 组件名称 (Component)  : FB_DL_CylStrokeTimeBank
 * 所属子库 (Sublibrary) : DL_Device
 * 当前版本 (Version)    : 1.0.0
 * 兼容性 (Platform)     : CODESYS 3.5+ / TwinCAT 3 / 汇川 InoProShop / 施耐德 Machine Expert
 *                         仅依赖 Standard.library（R_TRIG），零厂商私有库
 * 功能描述 (Function)   : 气缸行程时间分档趋势库。多缸（1..8）各自的行程完成
 *                         事件（bStrokeDone 沿 + nCylId + fStrokeTimeS）逐拍
 *                         建档：每缸记录 count/last/avg/min/max，并与基准时间
 *                         fBaseTimeS 比对输出劣化分档 eClass（0 正常 / 1 关注
 *                         / 2 预警 / 3 劣化），分档按最近耗时相对基准的劣化比
 *                         r = last/base 判定。维护性预测、气缸寿命台账场景。
 * 来源标签 (Origin)     : 自研线（IEC 61131-3 标准语义的道莅防御性实现，clean-room）
 * 边界语义 (Boundary)   : ① 缸号闸：nCylId 落于 1..8 域外 → 本拍拒收建档并
 *                         nWarnCnt 递增（信息级，不置故障级）；
 *                         ② 行程时间闸：fStrokeTimeS <= eps 或 NaN → 拒收
 *                         （传感器坏值不污染台账）；
 *                         ③ 劣化比除零防御：fBaseTimeS <= eps → 组态故障锁存
 *                         （分档判据整体失效必须可观测，R28 组态域闸覆盖）；
 *                         ④ 监视型事件建档，无主状态机（R23 公约）。
 * 输出语义 (Fallback)   : 【R191】bError = TRUE（组态故障）时全部建档动作冻结，
 *                         既有台账保持（不清零——台账是资产）；分档输出保持末值。
 * 码位     (Codes)      : 按 R297 范式零 16# 码位硬编码；错误出口 BOOL(bError)，
 *                         码位待主控收口统一派号。
 * 红线自检 (Redline)    : 7 项红线已自检：R1 零全局 ✓｜R2 零物理地址 ✓｜R3 纯 IEC ✓
 *                         R4 除零（基准 eps 闸）/下标钳位/NaN 拒收 ✓
 *                         R5 双语同行注释 ✓｜R6 N/A（监视型无状态机）✓
 *                         R7 R_TRIG 段 0 无条件刷新 ✓
 * 验收向量 (Acceptance) : V1 基准 1.0s，缸 3 上报 1.0s → r=1.0 → eClass[3]=0 正常；
 *                         V2 缸 3 上报 1.35s → r=1.35 → eClass[3]=1 关注；
 *                         V3 缸 3 上报 1.8s → eClass[3]=2 预警；2.6s → 3 劣化；
 *                         V4 缸号 0/9 → 拒收且 nWarnCnt 递增。
 * 修订历史 (Revision)   : 2026-11-20  v1.0.0  R49 首版（批 2 · 序号 9）
 *==============================================================================*)
TYPE E_DL_CstClass :
(
    eNormal   := 0,                          (* 正常：劣化比 < 1.2 / Normal: ratio < 1.2 *)
    eWatch    := 1,                          (* 关注：1.2 <= r < 1.5 / Watch band *)
    eWarning  := 2,                          (* 预警：1.5 <= r < 2.5 / Warning band *)
    eDegraded := 3                           (* 劣化：r >= 2.5 / Degraded band *)
);
END_TYPE

FUNCTION_BLOCK FB_DL_CylStrokeTimeBank
VAR_INPUT
    bStrokeDone : BOOL := FALSE;             (* 行程完成事件电平（内部取沿）[-] / Stroke-done event level *)
    nCylId      : INT := 1;                  (* 气缸编号，域 1..8，域外拒收 [缸] / Cylinder id, domain 1..8 *)
    fStrokeTimeS: LREAL := 0.0;              (* 本次行程耗时 [s] / Stroke time this event *)
    fBaseTimeS  : LREAL := 1.0;              (* 基准行程时间（分档分母），域 > eps [s] / Baseline stroke time *)
    bEnable     : BOOL := TRUE;              (* 建档使能，FALSE 时冻结不动台账 [-] / Enable *)
    bReset      : BOOL := FALSE;             (* 复位命令，上升沿清全部台账与告警 [-] / Reset command *)
END_VAR
VAR_OUTPUT
    aCnt    : ARRAY[1..8] OF DINT;           (* 各缸建档样本数 [个] / Sample count per cylinder *)
    aLast   : ARRAY[1..8] OF LREAL;          (* 各缸最近行程耗时 [s] / Last stroke time per cylinder *)
    aAvg    : ARRAY[1..8] OF LREAL;          (* 各缸平均行程耗时 [s] / Average per cylinder *)
    aMin    : ARRAY[1..8] OF LREAL;          (* 各缸最小行程耗时 [s] / Minimum per cylinder *)
    aMax    : ARRAY[1..8] OF LREAL;          (* 各缸最大行程耗时 [s] / Maximum per cylinder *)
    aeClass : ARRAY[1..8] OF E_DL_CstClass; (* 各缸劣化分档（按最近耗时相对基准）[-] / Class per cylinder *)
    bBanked : BOOL;                          (* 本拍完成一次建档的单拍脉冲 [-] / Bank-update single-scan pulse *)
    nWarnCnt: UDINT;                         (* 非法缸号/坏值拒收累计（信息级台账）[次] / Rejection counter *)
    bError  : BOOL;                          (* 组态故障锁存标志（基准时间非法）[-] / Config fault flag *)
END_VAR
VAR
    rtDone   : R_TRIG;                       (* 行程完成沿实例，段 0 无条件调用 / Stroke-done edge instance *)
    rtReset  : R_TRIG;                       (* 复位沿实例，段 0 无条件调用 / Reset edge instance *)
    _nId     : INT;                          (* 防御后生效缸号 [缸] / Sanitized cylinder id *)
    _bReject : BOOL;                         (* 本拍拒收当拍量（坏值/非法号）[-] / Reject this scan *)
    _fRatio  : LREAL;                        (* 劣化比 = last/base [-] / Degradation ratio *)
    _bFault  : BOOL;                         (* 组态故障锁存位 / Config fault latch bit *)
    _i       : INT;                          (* 复位清档游标 [-] / Reset clear cursor *)
END_VAR
VAR CONSTANT
    DL_CST_EPS   : LREAL := 1.0E-6;          (* 行程时间判零容差 [s] / Stroke time epsilon *)
    DL_CST_NMAX  : INT   := 8;               (* 缸容量上限 [缸] / Cylinder capacity limit *)
    DL_CST_DMAX  : DINT  := 1073741824;      (* 计数饱和上限 2^30（防回绕）[个] / Count saturation limit *)
    DL_CST_SUMMAX: LREAL := 1.0E15;          (* 均值递推饱和上限（防精度坍缩）[s] / Mean recursion saturation *)
    DL_R_WATCH   : LREAL := 1.2;             (* 关注档劣化比门限 [-] / Watch band ratio *)
    DL_R_WARNING : LREAL := 1.5;             (* 预警档劣化比门限 [-] / Warning band ratio *)
    DL_R_DEGRADE : LREAL := 2.5;             (* 劣化档劣化比门限 [-] / Degraded band ratio *)
END_VAR

(* —— 段 0：沿实例无条件刷新（R228A） —— *)
rtDone(CLK := bStrokeDone);                  (* 行程完成沿每拍必调 / Stroke edge every scan *)
rtReset(CLK := bReset);                      (* 复位沿每拍必调 / Reset edge every scan *)

(* —— 段 1：单拍量预清零（R107） —— *)
bBanked := FALSE;                            (* 建档单拍位预清，唯一分支置位 / Bank pulse preset *)
_bReject := FALSE;                           (* 拒收当拍量预清 / Reject preset *)

(* —— 段 2：组态闸故障锁存（分档分母失效必须可观测，R28 组态域闸；锁存至复位沿，R189） —— *)
IF (fBaseTimeS <= DL_CST_EPS) OR (fBaseTimeS <> fBaseTimeS) OR ((fBaseTimeS - fBaseTimeS) <> (fBaseTimeS - fBaseTimeS)) THEN
    _bFault := TRUE;                         (* 基准时间非法/非有限 → 锁存 / Illegal baseline, latch *)
END_IF

(* —— 段 3：复位沿处理（作用域：清故障 + 清全部缸档位 + 清告警台账，R283 逐项声明） —— *)
IF rtReset.Q THEN
    _bFault := FALSE;                        (* 清故障锁存 / Clear fault *)
    nWarnCnt := 0;                           (* 清拒收台账 / Clear counter *)
    _i := 1;                                 (* 游标起头重置（R227） / Cursor reset *)
    WHILE _i <= DL_CST_NMAX DO               (* 全缸档位清零（上电回夹防线） / Clear all banks *)
        aCnt[_i] := 0;                       (* 清计数 / Clear count *)
        aLast[_i] := 0.0;                    (* 清最近值 / Clear last *)
        aAvg[_i] := 0.0;                     (* 清均值 / Clear avg *)
        aMin[_i] := 0.0;                     (* 清最小值 / Clear min *)
        aMax[_i] := 0.0;                     (* 清最大值 / Clear max *)
        aeClass[_i] := E_DL_CstClass.eNormal;   (* 分档回归正常 / Class back to normal *)
        _i := _i + 1;                        (* 游标递进 / Cursor advance *)
    END_WHILE
END_IF

(* —— 段 4：建档事件处理（监视型纯派生，无 CASE 相；使能与组态双闸） —— *)
IF rtDone.Q AND bEnable AND NOT _bFault THEN
    _nId := nCylId;                          (* 生效缸号初值 / Id init *)
    IF (_nId < 1) OR (_nId > DL_CST_NMAX) THEN
        _bReject := TRUE;                    (* 非法缸号拒收 / Illegal id reject *)
    END_IF
    IF (fStrokeTimeS <= DL_CST_EPS) OR (fStrokeTimeS <> fStrokeTimeS) OR ((fStrokeTimeS - fStrokeTimeS) <> (fStrokeTimeS - fStrokeTimeS)) THEN
        _bReject := TRUE;                    (* 坏值/NaN 拒收（不污染台账） / Bad value reject *)
    END_IF
    IF _bReject THEN
        nWarnCnt := nWarnCnt + 1;            (* 信息级台账递增（不置 bError，R90 口径） / Info counter, not fault *)
    ELSE
        aLast[_nId] := fStrokeTimeS;         (* 记最近耗时 / Store last *)
        IF aCnt[_nId] < DL_CST_DMAX THEN
            aAvg[_nId] := (aAvg[_nId] * DINT_TO_LREAL(aCnt[_nId]) + fStrokeTimeS) / DINT_TO_LREAL(aCnt[_nId] + 1);   (* 增量均值，除子恒 >= 1 / Incremental mean, divisor >= 1 *)
            aCnt[_nId] := aCnt[_nId] + 1;    (* 计数递增（回绕防护） / Count advance *)
        END_IF
        IF (aMin[_nId] <= 0.0) OR (fStrokeTimeS < aMin[_nId]) THEN
            aMin[_nId] := fStrokeTimeS;      (* 最小值更新 / Min update *)
        END_IF
        IF fStrokeTimeS > aMax[_nId] THEN
            aMax[_nId] := fStrokeTimeS;      (* 最大值更新 / Max update *)
        END_IF
        _fRatio := fStrokeTimeS / fBaseTimeS;   (* 劣化比：分母已过组态闸，无除零 / Ratio, baseline gated *)
        IF _fRatio >= DL_R_DEGRADE THEN
            aeClass[_nId] := E_DL_CstClass.eDegraded;   (* 劣化档 / Degraded *)
        ELSIF _fRatio >= DL_R_WARNING THEN
            aeClass[_nId] := E_DL_CstClass.eWarning;    (* 预警档 / Warning *)
        ELSIF _fRatio >= DL_R_WATCH THEN
            aeClass[_nId] := E_DL_CstClass.eWatch;      (* 关注档 / Watch *)
        ELSE
            aeClass[_nId] := E_DL_CstClass.eNormal;     (* 正常档（IF 链带 ELSE 兜底，R285） / Normal *)
        END_IF
        bBanked := TRUE;                     (* 建档单拍脉冲 / Bank pulse *)
    END_IF
END_IF

(* —— 段 5：出口映射（R191 名实同源） —— *)
bError := _bFault;                           (* 组态故障镜像 / Config fault mirror *)
END_FUNCTION_BLOCK

(* ---- FB_DL_DamperBitDiag.st ---- *)
(*
  FB_DL_DamperBitDiag  —  风阀执行器位诊断打包/解包（位段提取 + 位打包复用） / Damper actuator bit diagnostics pack/unpack: field extraction and packing reuse
  分类 Category : DL_Device
  版本 Version  : 1.0.0
  来源 Source   : t2-1-lgf-bitlogic — 位逻辑族深化（与 AhuDamperStuckDiag 卡滞诊断/FreshAirStepperDamper 步进执行器分工：本件为状态字位诊断打包件）
  溯源 Origin   : clean-room 实现，未复制任何源码行
  功能 Function : 1) 位段解包：uStatusWord 固定位段提取——位 0 开限位、位 1 关限位、
                  位 2 运行位（掩码 AND 提取，移位量仅常量 0/1，R48 合规）；
                  2) 位打包复用：uDiagWord 输出按固定布局重打包（位 0..2 原样
                  直通、位 8 关键故障锁存镜像、位 9 反馈矛盾锁存镜像），
                  打包与解包同件承载（复用声明）；
                  3) 关键故障位检出：uStatusWord AND uFaultMask ≠ 0
                  → 0525 锁存（掩码域闸 uFaultMask ≠ 0）；
                  4) 反馈矛盾：开限与关限同 TRUE 持续 tContraWin → 0526 锁存
                  （R190 归因唯一：关键故障走 0525，矛盾走 0526）；
                  5) 故障级：0525 关键故障位锁存 / 0526 限位反馈矛盾锁存 /
                  0527 组态非法（掩码空）+ ELSE 兜底归并；
                  6) 信息级三码：诊断位检出 / 打包字更新 / 诊断复位（单拍沿）；
                  7) 解除式全当拍量（R240 落地），逐 BOOL 标注见段 4。
  边界 Boundary : ① 分段理由（R192）：段 0003 故障带 03A0~03FF 于 R42 用尽，
                  启用 05xx 副带续编，避开 0590~0599 判错位段；
                  ② 位段覆盖声明：本件仅校验位 0..2 与 uFaultMask 交叠域，
                  位 3..7/10..15 不做校验（域外是「不存在」而非「非法」，R57 口径）；
                  ③ 打包字位 8/9 为锁存镜像派生式（R28 建议位派生口径）；
                  ④ 无 GVL 依赖：纯引脚输入输出，无外部变量引用，无物理 IO 地址。
  依赖 Depends  : Standard.library（TON / R_TRIG）
  码表 Error codes（Device 段 0003，窗口 0525~0527 / 042B~042D）:
    16#0003_0525 故障级：关键故障位检出锁存（uFaultMask 交叠非零），锁存至 bReset
    16#0003_0526 故障级：限位反馈矛盾锁存（开限与关限同 TRUE 持续 tContraWin），锁存至 bReset
    16#0003_0527 故障级：组态非法（uFaultMask = 0）或相位落 ELSE 兜底（归并声明），锁存至 bReset
    16#0003_042B 信息级：诊断位检出沿（关键位或矛盾位首次置位拍）
    16#0003_042C 信息级：打包字更新沿（uDiagWord 与上拍不同拍）
    16#0003_042D 信息级：诊断复位沿（bDiagRst 生效拍）
  修订历史 Revision :
    2026-11-19  v1.0.0  R42 首版（批次 4 · 序号 4）
*)

TYPE E_DL_DbdState :
(
    eIdle  := 0,     // 待命：打包字静态承载 / Idle, packed word steady
    eDiag  := 10,    // 诊断中：位判据承载 / Diag, bit verdicts engaged
    eFault := 90     // 故障：关键位或矛盾锁定 / Fault, latched
);
END_TYPE

FUNCTION_BLOCK FB_DL_DamperBitDiag
VAR_INPUT
    uStatusWord  : WORD := 16#0000;   // 执行器状态字（位 0 开限/位 1 关限/位 2 运行）[-] / Actuator status word
    uFaultMask   : WORD := 16#0008;   // 关键故障位掩码（位 3 默认），域 ≠ 0 / Key fault bit mask
    tContraWin   : TIME := T#500MS;   // 反馈矛盾确认窗 [ms]，域 > 0 / Feedback contradiction window
    bDiagEn      : BOOL := FALSE;     // 诊断使能（电平）[-] / Diag enable, level
    bDiagRst     : BOOL := FALSE;     // 诊断复位指令，上升沿清锁存与打包镜像 [-] / Diag reset command edge
    bReset       : BOOL := FALSE;     // 复位，上升沿清故障锁存 / Reset edge clears fault latch
END_VAR
VAR_OUTPUT
    eState       : E_DL_DbdState;     // 状态出口，段尾单点映射 / State outlet
    uDiagWord    : WORD;              // 诊断打包字（固定布局见头注释）/ Diagnostic packed word
    bLimOpen     : BOOL;              // 开限位解包出口（位 0）[-] / Limit-open unpacked outlet
    bLimClosed   : BOOL;              // 关限位解包出口（位 1）[-] / Limit-closed unpacked outlet
    bRunning     : BOOL;              // 运行位解包出口（位 2）[-] / Running unpacked outlet
    bError       : BOOL;              // 故障锁存标志 / Fault latch flag
    nErrId       : UDINT;             // 事件码，0 = 无事件 / Event code
END_VAR
VAR
    tonContra    : TON;               // 反馈矛盾确认窗（电平式），无条件刷新 / Contradiction timer
    _eState      : E_DL_DbdState := E_DL_DbdState.eIdle;  // 内部相位（CASE 唯一写入目标，初值安全侧）/ Internal phase, safe init
    rtDiagRst    : R_TRIG;            // 诊断复位沿实例，无条件刷新 / Diag reset edge instance
    rtReset      : R_TRIG;            // 复位沿实例，无条件刷新 / Reset edge instance
    _bLimOpen    : BOOL;              // 开限位当拍量（掩码提取）[-] / Limit-open current-scan flag
    _bLimClosed  : BOOL;              // 关限位当拍量（掩码提取）[-] / Limit-closed current-scan flag
    _bRunning    : BOOL;              // 运行位当拍量（掩码提取）[-] / Running current-scan flag
    _bKeyFault   : BOOL;              // 关键故障位当拍量（掩码交叠）[-] / Key-fault bit flag
    _bContra     : BOOL;              // 限位矛盾当拍量 [-] / Limit contradiction flag
    _uDiagPrev   : WORD;              // 上拍打包字镜像（更新沿判据）/ Previous packed word mirror
    _bFault      : BOOL;              // 故障锁存位（锁存量）/ Latched fault bit
    _uFault      : UDINT;             // 故障码锁存（锁存量）/ Latched fault code
    _uInfo       : UDINT;             // 信息码，每拍重算 / Transient info code
END_VAR

(* —— 段 0：定时器与沿实例无条件周期刷新（禁置于 IF/CASE 内） —— *)
_bLimOpen   := (uStatusWord AND 16#0001) <> WORD#0;  // 位 0 开限（掩码提取，当拍量）
_bLimClosed := (uStatusWord AND 16#0002) <> WORD#0;  // 位 1 关限（掩码提取，当拍量）
_bRunning   := (uStatusWord AND 16#0004) <> WORD#0;  // 位 2 运行（掩码提取，当拍量）
_bKeyFault  := (uStatusWord AND uFaultMask) <> WORD#0;   // 关键故障位交叠（当拍量）
_bContra    := _bLimOpen AND _bLimClosed;            // 限位矛盾（当拍量）
rtDiagRst(CLK := bDiagRst);          // 诊断复位沿（每拍必调）
rtReset(CLK := bReset);              // 复位沿（每拍必调）
tonContra(IN := bDiagEn AND _bContra, PT := tContraWin); // 矛盾窗（电平式，矛盾消失自动断 IN）

(* —— 段 1：单拍量预清零（锁存量 _bFault/_uFault 不入清单，禁同拍抹除） —— *)
_uInfo := 16#0000_0000;             // 信息码每拍重算
nErrId := 16#0000_0000;             // 事件码缺省无事件

(* —— 段 2：复位沿 + 组态域闸（判据当拍量） —— *)
IF rtReset.Q THEN                   // rtReset.Q = 当拍量
    _bFault := FALSE;               // 清故障锁存位
    _uFault := 16#0000_0000;        // 清故障锁存码
END_IF
IF uFaultMask = WORD#0 THEN         // 掩码域闸（WORD 判等合规）
    _uFault := 16#0003_0527;        // 故障级：组态非法
    _bFault := TRUE;                // 故障标志与码位配对（R45）
END_IF
IF rtDiagRst.Q THEN                 // 诊断复位沿（当拍量）
    uDiagWord := WORD#0;            // 打包字清零
    _uDiagPrev := WORD#0;           // 镜像同步清零
    _uInfo := 16#0003_042D;         // 信息级：诊断复位沿
END_IF

(* —— 段 3：关键位与矛盾锁存（判据当拍量/电平式窗） —— *)
IF (NOT _bFault) AND bDiagEn AND _bKeyFault THEN
    _uFault := 16#0003_0525;        // 故障级：关键故障位锁存
    _bFault := TRUE;
    _uInfo := 16#0003_042B;         // 信息级：诊断位检出沿
END_IF
IF (NOT _bFault) AND tonContra.Q THEN
    _uFault := 16#0003_0526;        // 故障级：限位反馈矛盾锁存
    _bFault := TRUE;
    _uInfo := 16#0003_042B;         // 信息级：诊断位检出沿（同检出口，成因由 nErrId 区分声明）
END_IF

(* —— 段 4：故障解除式（R240 落地，逐 BOOL 标注）：
     rtReset.Q = 当拍量；rtDiagRst.Q = 当拍量；NOT _bKeyFault = 当拍量；
     NOT _bContra = 当拍量；NOT bDiagEn = 当拍量。均不含锁存量（_bFault/_uFault），
     解除边真实可达（状态字恢复 + 复位/诊断复位沿）。 —— *)
IF (rtReset.Q OR rtDiagRst.Q) AND (NOT _bKeyFault) AND (NOT _bContra) THEN
    _bFault := FALSE;               // 清故障锁存位（锁存量，仅此当拍量解除沿可清）
    _uFault := 16#0000_0000;        // 清故障锁存码（锁存量，仅本当拍量解除沿可清）
    IF _eState = E_DL_DbdState.eFault THEN
        _eState := E_DL_DbdState.eIdle;     // 故障相迁出：回待命
    END_IF
END_IF

(* —— 段 5：相位机（CASE 全覆盖 + ELSE 兜底） —— *)
CASE _eState OF

E_DL_DbdState.eIdle:
    IF bDiagEn AND (NOT _bFault) THEN
        _eState := E_DL_DbdState.eDiag;     // 使能：进诊断相
    END_IF

E_DL_DbdState.eDiag:
    IF NOT bDiagEn THEN
        _eState := E_DL_DbdState.eIdle;     // 撤使能：回待命相
    END_IF
    (* 关键位/矛盾迁出在段 3 承载 *)

E_DL_DbdState.eFault:
    ;                               // 故障相：锁存码回放，等解除沿（段 4 承载迁出）

ELSE
    _uFault := 16#0003_0527;        // 故障级：非法相位兜底（归并组态码，码表声明）
    _bFault := TRUE;
    _eState := E_DL_DbdState.eFault;    // 强制回故障相

END_CASE

(* —— 段 6：位打包（固定布局：位 0..2 直通、位 8/9 锁存镜像派生，R28 派生口径） —— *)
uDiagWord := WORD#0;                // 打包字每拍重构（位段固定，无残留位）
IF _bLimOpen THEN
    uDiagWord := uDiagWord OR 16#0001;      // 位 0 直通
END_IF
IF _bLimClosed THEN
    uDiagWord := uDiagWord OR 16#0002;      // 位 1 直通
END_IF
IF _bRunning THEN
    uDiagWord := uDiagWord OR 16#0004;      // 位 2 直通
END_IF
IF _bFault THEN
    uDiagWord := uDiagWord OR 16#0100;      // 位 8：故障锁存镜像（派生式）
END_IF
IF _uFault = 16#0003_0526 THEN      // 矛盾码判等（UDINT 合规）
    uDiagWord := uDiagWord OR 16#0200;      // 位 9：矛盾锁存镜像（派生式）
END_IF
IF uDiagWord <> _uDiagPrev THEN     // 更新沿（当拍量判据）
    _uInfo := 16#0003_042C;         // 信息级：打包字更新沿
END_IF
_uDiagPrev := uDiagWord;            // 更新沿判据快照（段末统一写）

(* —— 段 7：出口单点映射（名实同源；锁存码回放，禁同拍抹除） —— *)
IF _bFault THEN
    nErrId := _uFault;              // 故障锁存码回放
ELSE
    nErrId := _uInfo;               // 信息码
END_IF
bError := _bFault;                  // 故障标志与锁存位同源
bLimOpen := _bLimOpen;              // 解包出口（当拍量直出）
bLimClosed := _bLimClosed;          // 解包出口（当拍量直出）
bRunning := _bRunning;              // 解包出口（当拍量直出）
eState := _eState;                  // 状态出口单点映射

END_FUNCTION_BLOCK

(* ---- FB_DL_DateCoderSync.st ---- *)
(*==============================================================================
 * 组件名称 (Component)  : FB_DL_DateCoderSync
 * 所属子库 (Sublibrary) : DL_Device
 * 当前版本 (Version)    : 1.0.0
 * 兼容性 (Platform)     : CODESYS 3.5 / TwinCAT 3 / 汇川 InoProShop / Machine Expert
 *                         仅依赖纯 IEC 61131-3 标准元素，零厂商方言
 * 功能描述 (Function)   : 喷码/打码同步：R_TRIG 采编码器脉冲 → 计数器带偏移
 *                         → 计满修正分频比触发一拍喷印（TP 成形脉宽）；产品检测
 *                         丢失超时 → 跳过本袋并计数；偏移限幅后合成目标（以
 *                         >= 比较替代取模，杜绝负余数）；相位诊断委托 FC_DL_ModPos。
 * 溯源 (Origin)         : 道莅 clean-room 防御性实现
 * 本文件内含 (Contains) : TYPE E_DL_CoderErr / FUNCTION_BLOCK FB_DL_DateCoderSync
 * 依赖 (Depends)        : DL_MathData/FC_DL_ModPos
 * 红线自检 (Redline)    : 无外部全局变量、无硬件地址直引 ｜ 全变量中英双语同行注释
 *                         分频比下限钳 1 防除零 ｜ 偏移双向限幅 ｜ 枚举成员全部显式赋值
 *                         R_TRIG/TP/TON 实例每周期无条件调用（仅输入条件化）｜
 *                         负余数防御：目标合成用 >= 比较，不裸用取模
 * 错误码表 (Codes)      : 16#0003_039D 就绪
 *                         16#0003_039E 信息级 分频比非法(已钳 1)
 *                         16#0003_039F 信息级 偏移越界(已钳制)
 *                         16#0003_03A0 信息级 产品信号超时(已跳过)
 *                         16#0003_03A1 信息级 正常喷印中
 * 修订历史 (Revision)   : 2026-11-17  v1.0.0  首版入库 · R27 · 阶段三批 2
 * 验收向量 (Acceptance) : 分频 10，偏移 0：第 10 个编码脉冲 → bPrintTrig 一拍脉宽；
 *                         偏移 +3 → 第 13 个脉冲触发；分频 0 → 钳 1 且 039E；
 *                         产品信号丢失超 tProdMax → 跳过且 03A0
 *============================================================================*)

(*-----------------------------------------------------------------------------
 * 枚举: E_DL_CoderErr（归属 DL_Device，与 FB_DL_DateCoderSync 同文件）
 *----------------------------------------------------------------------------*)
TYPE E_DL_CoderErr :
(
    eReady      := 16#0003_039D,   // 就绪 / Ready
    eDivClamped := 16#0003_039E,   // 信息级：分频比非法已钳 1 / Info: division ratio clamped to 1
    eOffsetClamp:= 16#0003_039F,   // 信息级：偏移越界已钳制 / Info: offset clamped
    eProdSkip   := 16#0003_03A0,   // 信息级：产品信号超时已跳过 / Info: product timeout, skipped
    ePrinting   := 16#0003_03A1    // 信息级：正常喷印中 / Info: printing active
);
END_TYPE

(*==============================================================================
 * 功能块: FB_DL_DateCoderSync
 * 调用约定: 每个扫描周期无条件调用一次。
 *============================================================================*)
FUNCTION_BLOCK FB_DL_DateCoderSync
VAR_INPUT
    bEncoderPulse  : BOOL;             // 编码器脉冲输入 / Encoder pulse input
    uDivRatio      : UINT;             // 分频比 [脉冲每触发]，有效域 1~10000 / Division ratio [pulses per trigger]
    nOffsetCounts  : DINT;             // 偏移补偿 [脉冲]，有效域 -1000~1000 / Offset compensation [pulses]
    bProductDetect : BOOL;             // 产品到位信号 / Product present signal
    tPulseWidth    : TIME := T#10MS;   // 喷印触发脉宽 [毫秒] / Print trigger pulse width [ms]
    tProdMax       : TIME := T#5S;     // 产品信号丢失超时 [秒] / Product signal timeout [s]
END_VAR
VAR_OUTPUT
    bPrintTrig     : BOOL;             // 喷印触发（TP 成形脉宽）/ Print trigger, TP-formed pulse
    uPulseCount    : UDINT;            // 累计编码脉冲 [个]，诊断 / Accumulated pulse count [pcs]
    uSkipCount     : UDINT;            // 跳过计数 [次]，诊断 / Skipped-product count [pcs]
    nPhaseDiag     : DINT;             // 相位诊断（当前计数对目标取正余数）/ Phase diagnostic, positive remainder
    eErr           : E_DL_CoderErr;    // 错误码 / Error code
END_VAR
VAR
    fbEncTrig      : R_TRIG;           // 编码脉冲上升沿实例（无条件调用）/ Encoder pulse edge instance
    fbPrintPulse   : TP;               // 喷印脉宽定时器实例（无条件调用）/ Print pulse timer instance
    bTrigReq       : BOOL;             // 触发请求锁存（TP 输入条件源）/ Trigger request latch, TP input source
    tonProdLost    : TON;              // 产品信号丢失计时器（无条件调用）/ Product-lost timer
    nCount         : DINT;             // 本袋脉冲计数 [个] / Pulse count for the current bag [pcs]
    nTarget        : DINT;             // 合成触发目标（分频+偏移，下限 1）/ Composite trigger target [pulses]
    uDivUse        : UINT;             // 生效分频比（钳位后）[脉冲每触发] / Effective division ratio
    nOffsetUse     : DINT;             // 生效偏移（限幅后）[脉冲] / Effective offset [pulses]
    uPulseAcc      : UDINT;            // 累计脉冲工作副本（饱和自增）[个] / Accumulated pulse working copy [pcs]
    uSkipAcc       : UDINT;            // 跳过计数工作副本（饱和自增）[次] / Skip count working copy [pcs]
    uPhaseErr      : UDINT;            // 委托取模错误码（0 = 无错）/ Delegate modulo error id
END_VAR
VAR CONSTANT
    DL_COD_DIV_MAX    : UINT := 10000;          // 分频比上限 [脉冲每触发] / Division ratio upper bound
    DL_COD_OFF_MIN    : DINT := -1000;          // 偏移下限 [脉冲] / Offset lower bound [pulses]
    DL_COD_OFF_MAX    : DINT := 1000;           // 偏移上限 [脉冲] / Offset upper bound [pulses]
    DL_COD_TARGET_MIN : DINT := 1;              // 触发目标下限 [脉冲]（防除零与零目标死锁）/ Target lower bound [pulses]
    DL_COD_CNT_SAT    : UDINT := 16#FFFF_FFFE;  // 累计计数饱和值 [个] / Count saturation [pcs]
END_VAR

(*------------------------------------------------------------------------------
 * 段 1｜沿检测/TP/TON 实例每周期无条件调用（仅输入条件化）
 *----------------------------------------------------------------------------*)
fbEncTrig(CLK := bEncoderPulse);                      // 编码脉冲沿检测无条件刷新 / encoder edge refreshed unconditionally
fbPrintPulse(IN := bTrigReq AND bProductDetect, PT := tPulseWidth);   // 喷印脉宽成形（IN 条件化，请求锁存源）/ print pulse formed
tonProdLost(IN := NOT bProductDetect, PT := tProdMax);   // 产品信号丢失计时 / product-lost timing

(*------------------------------------------------------------------------------
 * 段 2｜分频比钳位（下限 1 防除零与零目标死锁）与偏移双向限幅
 *----------------------------------------------------------------------------*)
eErr := E_DL_CoderErr.eReady;                         // 预置就绪 / preset ready
uDivUse := uDivRatio;                                 // 分频工作副本 / division working copy
IF (uDivUse < 1) OR (uDivUse > DL_COD_DIV_MAX) THEN
    uDivUse := 1;                                     // 分频非法钳 1 / division clamped to 1
    eErr := E_DL_CoderErr.eDivClamped;                // 信息级：分频比非法 / info: ratio clamped
END_IF
nOffsetUse := nOffsetCounts;                          // 偏移工作副本 / offset working copy
IF nOffsetUse < DL_COD_OFF_MIN THEN
    nOffsetUse := DL_COD_OFF_MIN;                    // 偏移下限钳位 / offset floored
    IF eErr = E_DL_CoderErr.eReady THEN
        eErr := E_DL_CoderErr.eOffsetClamp;          // 信息级：偏移越界 / info: offset clamped
    END_IF
ELSIF nOffsetUse > DL_COD_OFF_MAX THEN
    nOffsetUse := DL_COD_OFF_MAX;                    // 偏移上限钳位 / offset capped
    IF eErr = E_DL_CoderErr.eReady THEN
        eErr := E_DL_CoderErr.eOffsetClamp;          // 信息级：偏移越界 / info: offset clamped
    END_IF
END_IF

(*------------------------------------------------------------------------------
 * 段 3｜合成触发目标：分频 + 偏移，下限 1；以 >= 比较替代取模，杜绝负余数
 *----------------------------------------------------------------------------*)
nTarget := UINT_TO_DINT(uDivUse) + nOffsetUse;        // 合成目标 [脉冲] / composite target [pulses]
IF nTarget < DL_COD_TARGET_MIN THEN
    nTarget := DL_COD_TARGET_MIN;                    // 目标下限钳位 / target floored
END_IF

(*------------------------------------------------------------------------------
 * 段 4｜产品信号丢失超时：跳过本袋计数并清计数器（信息级 03A0）
 *----------------------------------------------------------------------------*)
IF tonProdLost.Q THEN
    IF nCount > 0 THEN
        nCount := 0;                                 // 跳过本袋：计数清零 / skip bag: counter cleared
        IF uSkipAcc < DL_COD_CNT_SAT THEN
            uSkipAcc := uSkipAcc + 1;                // 跳过计数饱和自增 [次] / saturating skip increment
        END_IF
        IF eErr = E_DL_CoderErr.eReady THEN
            eErr := E_DL_CoderErr.eProdSkip;         // 信息级：产品信号超时 / info: product timeout
        END_IF
    END_IF
END_IF

(*------------------------------------------------------------------------------
 * 段 5｜编码脉冲计数与触发：计满合成目标即触发（TP 已在段 1 成形脉宽）
 *----------------------------------------------------------------------------*)
IF fbEncTrig.Q THEN
    nCount := nCount + 1;                            // 脉冲计数 [个] / pulse counted
    IF uPulseAcc < DL_COD_CNT_SAT THEN
        uPulseAcc := uPulseAcc + 1;                  // 累计脉冲饱和自增 [个] / saturating pulse increment
    END_IF
    IF nCount >= nTarget THEN
        bTrigReq := TRUE;                            // 触发请求锁存（TP 下拍成形脉宽）/ trigger request latched
        nCount := 0;                                 // 触发后计数清零 / counter cleared after trigger
    END_IF
END_IF
IF fbPrintPulse.Q THEN
    bTrigReq := FALSE;                               // 脉宽完成：请求解锁 / pulse done: request released
END_IF
bPrintTrig := fbPrintPulse.Q;                        // 喷印触发输出（TP 成形）/ print trigger output
IF bPrintTrig THEN
    IF eErr = E_DL_CoderErr.eReady THEN
        eErr := E_DL_CoderErr.ePrinting;             // 信息级：正常喷印中 / info: printing active
    END_IF
END_IF
uPulseCount := uPulseAcc;                            // 累计脉冲输出 [个] / accumulated pulse output
uSkipCount := uSkipAcc;                              // 跳过计数输出 [次] / skip count output

(*------------------------------------------------------------------------------
 * 段 6｜相位诊断：委托 FC_DL_ModPos 防负余数（计数为非负，防御仍委托）
 *----------------------------------------------------------------------------*)
nPhaseDiag := FC_DL_ModPos(nValue := nCount, nModulus := nTarget, eErr => uPhaseErr);   // 正余数诊断 [个] / positive-remainder diagnostic
IF uPhaseErr <> 0 THEN
    nPhaseDiag := 0;                                 // 委托异常诊断归零 / diagnostic zeroed on delegate error
END_IF
END_FUNCTION_BLOCK

(* ---- FB_DL_DeviceHealthArbiter.st ---- *)
(*
    FB_DL_DeviceHealthArbiter —— NE107 多源健康聚合仲裁
    ------------------------------------------------------------------
    分类      : DL_Device / Diagnostics
    前缀      : FB_DL_
    版本      : 1.0.0
    溯源      : NAMUR NE107 公开的六态健康语言（只借六态语义与「编号即仲裁优先级」的
                组织事实，不复制任何条款文本）；聚合算法、分级位图、首出三律、错误分级与
                码位 100% 自有；E_DL_Ne107Status 的唯一属主为 I_DL_DeviceHealth，
                本件只引用不重声明（R70 全库唯一断言）；
                clean-room 重写，未复制任何闭源厂商源码
    平台      : 纯 IEC 61131-3，CODESYS V3.5+ / TwinCAT 3 / InoProShop 通用
    作者      : 道莅代码库 · PLC编程专家（R19）
    ------------------------------------------------------------------
    功能说明  : 把 N 路设备健康态（阀 / 电机 / 仪表 / 变频器）聚合成一个整机健康结论，
                并回答现场两个必答题：「现在最严重的是哪一类」与「是谁先报的」。
                核心防御：① 仲裁次序 = 枚举编号（eFailure 0 < eCheckFunction 10 <
                   eMaintenanceReq 20 < eOutOfSpec 30 < eOk 40 < eUnknown 99），
                   本件不自造第二套优先级（同族纪律）；
                ② Unknown 不遮蔽：只要有任一源为已知且非 OK 态，聚合结论就不得为
                   eUnknown——现场最常见的误判是一路通道没配好导致整机显示「未知」，
                   把真故障压掉；
                ③ 首出仅锁存一次，复位沿在仲裁之后生效且当拍不重新锁存；
                ④ 平台越界写入的非法枚举值落 ELSE 分支归 eUnknown 并置故障级 0331；
                ⑤ 源数量越界时不索引任何数组，聚合结论回 eUnknown。
                职责边界：单源健康判定归各设备件，本件只做聚合与仲裁；PN 通道诊断聚合归
                FB_DL_ProfinetAlarmDiag，本件不吃协议细节。
    错误码    : 16#0003_016A 同拍多源同级别已按源索引最小仲裁 / 存在 Unknown 源但未遮蔽已知故障——信息级，正常防御
                16#0003_016B 预留禁用（信息级，不得挪用）
                16#0003_0330 源数量越界（不在 1~16）——故障级，聚合结论置 eUnknown 且不索引数组
                16#0003_0331 健康枚举值非法（CASE 落 ELSE）——故障级，该源按 eUnknown 处理并继续聚合
                16#0003_0332 预留禁用（故障级，不得挪用）
    码位总账  : 16#0003_016A 用 / 16#0003_016B 预留 ｜ 16#0003_0330 用 / 16#0003_0331 用 / 16#0003_0332 预留
    状态机    : R6 标注 N/A —— 本组件为纯函数无顺序状态机，无 CASE 可写，非法状态不可能出现
                （源态分派用的 CASE 是枚举映射表，不是顺序状态机，且含 ELSE 兜底）
    采样约定  : fbTrigReset 在本体首部无条件刷新；健康结论每拍实时刷新（不锁存），
                只有首出索引与通道锁存；与任务周期无关的纯组合仲裁。
    修订记录  : 2026-11-16 v1.0.0 首次入库（R19）
*)
FUNCTION_BLOCK FB_DL_DeviceHealthArbiter
VAR_INPUT
    bEnable            : BOOL;                // 使能，FALSE 输出 eUnknown 并冻结首出 / enable, FALSE outputs eUnknown and freezes the first-out
    bReset             : BOOL;                // 复位，上升沿清首出锁存（健康结论仍实时刷新）/ reset, rising edge clears the first-out latch, health stays live
    aeHealth           : ARRAY[0..15] OF E_DL_Ne107Status; // 各源健康态，枚举属主为 I_DL_DeviceHealth / source health states, owned by I_DL_DeviceHealth
    auChannelId        : ARRAY[0..15] OF UINT; // 各源对外通道号，可为 0 [通道] / external channel id per source, zero allowed [channel]
    uSrcCount          : UINT := 16;           // 有效源数 [路]，范围 1~16 / valid source count [ch], range 1~16
    bIncludeMaintenance : BOOL := TRUE;        // TRUE = 维护/校验类参与聚合，FALSE = 只聚 Failure / OutOfSpec / TRUE lets maintenance and check participate
END_VAR
VAR_OUTPUT
    eAggHealth         : E_DL_Ne107Status;     // 聚合后健康结论 / aggregated health conclusion
    uFirstIdx          : UINT;                // 首出源索引 0~15，无则 16#FFFF / first-out source index, sentinel 16#FFFF when none
    uFirstChannel      : UINT;                // 首出源对外通道号 [通道] / external channel id of the first-out source [channel]
    auLevelMask        : ARRAY[0..5] OF WORD;  // 分级位图，bit N = 源 N / level bitmap, bit N is source N
    uFaultSrcCount     : UINT;                // 处于 Failure 或 OutOfSpec 的源数 [路] / sources in Failure or OutOfSpec [ch]
    bDegraded          : BOOL;                // 存在维护/校验类但无故障类（可运行需处理）/ degraded, maintenance or check without a fault class
    eErr               : UDINT;               // 错误码，0=正常 / error id, 0=ok
    bError             : BOOL;                // 故障标志，eErr 为故障级时 TRUE / error flag, TRUE on fault-level eErr
END_VAR
VAR
    fbTrigReset        : R_TRIG;              // 复位上升沿实例，本体首部无条件刷新 / reset edge instance, refreshed unconditionally
    uIdx               : UINT;                // 源扫描游标 [路]，范围 0~15 / source scan cursor [ch], range 0~15
    uBucket            : UINT;                // 本源的位图分桶序号 [桶] / bitmap bucket index of this source [bucket]
    nRank              : INT;                 // 本源的仲裁等级（枚举编号）[无量纲] / arbitration rank of this source [dimensionless]
    nBestRank          : INT;                 // 已选出的最高优先级等级 [无量纲] / best rank selected so far [dimensionless]
    uBestIdx           : UINT;                // 已选出的首出候选索引 [路] / first-out candidate index [ch]
    bAnyKnown          : BOOL;                // 存在已知（非 Unknown）源 / at least one known source exists
    bAnyUnknown        : BOOL;                // 存在 Unknown 源 / at least one unknown source exists
    bAnyMaintain       : BOOL;                // 存在维护/校验类源 / at least one maintenance or check source exists
    bAnyFaultLevel     : BOOL;                // 存在故障类（Failure/OutOfSpec）源 / at least one fault class source exists
    bConsider          : BOOL;                // 本源参与聚合判定标志 / this source participates in the aggregation
    bIllegalEnum       : BOOL;                // 本拍出现非法枚举值 / an illegal enumeration value appeared in this cycle
    bFirstLatched      : BOOL;                // 首出已锁存 / first-out is latched
    uFirstInt          : UINT := 16#FFFF;     // 内部首出索引寄存，初值哨兵 / internal first-out index, initialised to the sentinel
    uFirstChInt        : UINT;                // 内部首出通道寄存 / internal first-out channel register
    bMultiSame         : BOOL;                // 同拍多源同级别 / multiple sources share the best rank this cycle
    uSameCnt           : UINT;                // 与最高优先级同级别的源数 [路] / sources sharing the best rank [ch]
    bInit              : BOOL := FALSE;       // 首扫标志，初值 FALSE，判据 NOT bInit / first-scan flag, initial FALSE, tested with NOT
END_VAR
VAR CONSTANT
    DL_HARB_SRC_MAX     : UINT := 16;         // 源数量上限 [路] / source count upper bound [ch]
    DL_HARB_NONE        : UINT := 16#FFFF;    // 无首出哨兵 [无量纲] / no first-out sentinel [dimensionless]
    DL_HARB_LEVELS      : UINT := 6;          // 分级桶数 [桶] / number of level buckets [bucket]
    DL_HARB_B_FAILURE   : UINT := 0;          // eFailure 桶号 [桶] / bucket index for eFailure
    DL_HARB_B_CHECK     : UINT := 1;          // eCheckFunction 桶号 [桶] / bucket index for eCheckFunction
    DL_HARB_B_MAINT     : UINT := 2;          // eMaintenanceReq 桶号 [桶] / bucket index for eMaintenanceReq
    DL_HARB_B_SPEC      : UINT := 3;          // eOutOfSpec 桶号 [桶] / bucket index for eOutOfSpec
    DL_HARB_B_OK        : UINT := 4;          // eOk 桶号 [桶] / bucket index for eOk
    DL_HARB_B_UNKNOWN   : UINT := 5;          // eUnknown 桶号 [桶] / bucket index for eUnknown
    DL_HARB_R_FAILURE   : INT := 0;           // eFailure 的仲裁等级（最严重）[无量纲] / rank of eFailure, the most severe
    DL_HARB_R_CHECK     : INT := 10;          // eCheckFunction 的仲裁等级 [无量纲] / rank of eCheckFunction
    DL_HARB_R_MAINT     : INT := 20;          // eMaintenanceReq 的仲裁等级 [无量纲] / rank of eMaintenanceReq
    DL_HARB_R_SPEC      : INT := 30;          // eOutOfSpec 的仲裁等级 [无量纲] / rank of eOutOfSpec
    DL_HARB_R_OK        : INT := 40;          // eOk 的仲裁等级 [无量纲] / rank of eOk
    DL_HARB_R_UNKNOWN   : INT := 99;          // eUnknown 的仲裁等级（不参与优先）[无量纲] / rank of eUnknown, excluded from priority
    DL_HARB_R_NONE      : INT := 100;         // 未选出任何等级的哨兵 [无量纲] / sentinel meaning no rank selected yet
    DL_HARB_BIT0        : WORD := 16#0001;    // 位图最低位掩码 [位图] / least significant bitmap mask [bitmap]
    DL_HARB_ZERO        : WORD := 16#0000;    // 位图零常量 [位图] / bitmap zero constant [bitmap]
    DL_HARB_CNT_ZERO    : UINT := 0;          // 无符号零常量 [无量纲] / unsigned zero constant [dimensionless]
END_VAR

// 段 1｜边沿实例无条件周期刷新（红线：严禁放入条件分支）/ segment 1, unconditional edge refresh
fbTrigReset(CLK := bReset);

// 段 2｜输出与中间量预置 / segment 2, preset outputs and intermediates
eAggHealth := eUnknown;                       // 缺省结论为未知 / default conclusion is unknown
uFirstIdx := DL_HARB_NONE;                    // 缺省无首出 / default no first-out
uFirstChannel := DL_HARB_CNT_ZERO;            // 缺省通道号 0 / default channel zero
uFaultSrcCount := DL_HARB_CNT_ZERO;           // 故障源计数清零 / clear the fault source count
bDegraded := FALSE;                           // 预置未降级 / preset not degraded
eErr := 0;                                    // 预置无错误 / preset no error
bError := FALSE;                              // 预置无故障 / preset no fault
bAnyKnown := FALSE;                           // 预置无已知源 / preset no known source
bAnyUnknown := FALSE;                         // 预置无未知源 / preset no unknown source
bAnyMaintain := FALSE;                        // 预置无维护类 / preset no maintenance source
bAnyFaultLevel := FALSE;                      // 预置无故障类 / preset no fault class source
nBestRank := DL_HARB_R_NONE;                  // 最高优先级哨兵 / best rank sentinel
uBestIdx := DL_HARB_NONE;                     // 首出候选哨兵 / first-out candidate sentinel
bIllegalEnum := FALSE;                        // 预置无非法枚举 / preset no illegal enumeration
uSameCnt := DL_HARB_CNT_ZERO;                 // 同级别计数清零 / clear the same-rank counter
FOR uIdx := 0 TO DL_HARB_LEVELS - 1 DO
    auLevelMask[uIdx] := DL_HARB_ZERO;        // 六个分级桶逐桶清零 / clear each of the six level buckets
END_FOR

// 段 3｜首扫初始化（唯一合法范式：初值 FALSE，判据 NOT bInit）/ segment 3, first-scan initialisation
IF NOT bInit THEN
    bFirstLatched := FALSE;                   // 首扫不留锁存 / no latch survives the first scan
    uFirstInt := DL_HARB_NONE;                // 首出索引回哨兵 / first-out index back to the sentinel
    uFirstChInt := DL_HARB_CNT_ZERO;          // 首出通道回 0 / first-out channel back to zero
    bInit := TRUE;                            // 首扫只做一次 / first scan runs once only
END_IF

// 段 4｜使能闸：失能输出未知并冻结首出（不索引数组）/ segment 4, enable gate
IF NOT bEnable THEN
    eAggHealth := eUnknown;                   // 失能即未知 / unknown while disabled
    uFirstIdx := uFirstInt;                   // 首出保持冻结 / the first-out stays frozen
    uFirstChannel := uFirstChInt;             // 通道保持冻结 / the channel stays frozen
    RETURN;                                   // 失能即出口 / disabled is the exit
END_IF

// 段 5｜源数量闸：越界即故障级，聚合结论回 eUnknown 且不索引数组 / segment 5, source count gate
IF (uSrcCount < 1) OR (uSrcCount > DL_HARB_SRC_MAX) THEN
    eErr := 16#0003_0330;                     // 源数量越界故障码 / source count out of range fault id
    bError := TRUE;                           // 置故障标志 / raise the error flag
    eAggHealth := eUnknown;                   // 结论回未知 / conclusion back to unknown
    RETURN;                                   // 故障级提前返回，不索引任何源 / early return, no source is indexed
END_IF

// 段 6｜逐源扫描：分桶、计故障类、选最高优先级、捕非法枚举 / segment 6, per source scan
FOR uIdx := 0 TO uSrcCount - 1 DO
    bConsider := TRUE;                        // 默认参与聚合 / participates by default
    CASE aeHealth[uIdx] OF
        eFailure:
            uBucket := DL_HARB_B_FAILURE;     // 落失效桶 / bucket for failure
            nRank := DL_HARB_R_FAILURE;       // 最严重等级 / the most severe rank
            bAnyKnown := TRUE;                // 已知态 / a known state
            bAnyFaultLevel := TRUE;           // 故障类 / fault class
            uFaultSrcCount := uFaultSrcCount + 1; // 故障源计数加一 / increment the fault source count
        eCheckFunction:
            uBucket := DL_HARB_B_CHECK;       // 落功能校验桶 / bucket for function check
            nRank := DL_HARB_R_CHECK;         // 校验等级 / check rank
            bAnyKnown := TRUE;                // 已知态 / a known state
            bAnyMaintain := TRUE;             // 维护/校验类 / maintenance or check class
        eMaintenanceReq:
            uBucket := DL_HARB_B_MAINT;       // 落维护桶 / bucket for maintenance required
            nRank := DL_HARB_R_MAINT;         // 维护等级 / maintenance rank
            bAnyKnown := TRUE;                // 已知态 / a known state
            bAnyMaintain := TRUE;             // 维护/校验类 / maintenance or check class
        eOutOfSpec:
            uBucket := DL_HARB_B_SPEC;        // 落超规格桶 / bucket for out of specification
            nRank := DL_HARB_R_SPEC;          // 超规格等级 / out of specification rank
            bAnyKnown := TRUE;                // 已知态 / a known state
            bAnyFaultLevel := TRUE;           // 故障类 / fault class
            uFaultSrcCount := uFaultSrcCount + 1; // 故障源计数加一 / increment the fault source count
        eOk:
            uBucket := DL_HARB_B_OK;          // 落正常桶 / bucket for OK
            nRank := DL_HARB_R_OK;            // 正常等级 / the OK rank
            bAnyKnown := TRUE;                // 已知态 / a known state
        eUnknown:
            uBucket := DL_HARB_B_UNKNOWN;     // 落未知桶 / bucket for unknown
            nRank := DL_HARB_R_UNKNOWN;       // 未知等级（不参与优先）/ unknown rank, excluded from priority
            bAnyUnknown := TRUE;              // 存在未知源 / an unknown source exists
            bConsider := FALSE;               // 未知源不参与聚合 / an unknown source never participates
        ELSE
            uBucket := DL_HARB_B_UNKNOWN;     // 非法枚举归未知桶（红线 4：ELSE 兜底）/ illegal values fall into the unknown bucket
            nRank := DL_HARB_R_UNKNOWN;       // 按未知等级处理 / treated as unknown rank
            bAnyUnknown := TRUE;              // 计入未知源 / counted as an unknown source
            bConsider := FALSE;               // 不参与聚合 / never participates
            bIllegalEnum := TRUE;             // 记录非法枚举 / remember the illegal enumeration
        END_CASE
    auLevelMask[uBucket] := auLevelMask[uBucket] OR SHL(DL_HARB_BIT0, uIdx); // 置位图，uIdx ≤ 15 移位安全 / set the bitmap bit, the shift never exceeds 15

    // 段 7｜聚合参与判定：维护类是否计入由调用方策略决定 / segment 7, participation policy
    IF bConsider AND (NOT bIncludeMaintenance) THEN
        IF (uBucket = DL_HARB_B_CHECK) OR (uBucket = DL_HARB_B_MAINT) THEN
            bConsider := FALSE;               // 策略禁止时维护/校验类不进聚合，但仍进位图 / excluded from the aggregation but still visible in the bitmap
        END_IF
    END_IF

    // 段 8｜最高优先级仲裁：等级更小者胜，同级取源索引最小 / segment 8, best rank arbitration
    IF bConsider AND (nRank < nBestRank) THEN
        nBestRank := nRank;                   // 记下新的最高优先级 / remember the new best rank
        uBestIdx := uIdx;                     // 记下首出候选索引 / remember the candidate index
        uSameCnt := 1;                        // 同级别计数复位 / reset the same-rank counter
    ELSIF bConsider AND (nRank = nBestRank) THEN
        uSameCnt := uSameCnt + 1;             // 同级别源计数 / count the sources sharing the rank
    END_IF
END_FOR

// 段 9｜等级回映射为枚举（含兜底，绝不返回未定义值）/ segment 9, rank to enumeration mapping
CASE nBestRank OF
    DL_HARB_R_FAILURE:
        eAggHealth := eFailure;               // 聚合结论：失效 / aggregated failure
    DL_HARB_R_CHECK:
        eAggHealth := eCheckFunction;         // 聚合结论：功能校验 / aggregated function check
    DL_HARB_R_MAINT:
        eAggHealth := eMaintenanceReq;        // 聚合结论：需要维护 / aggregated maintenance required
    DL_HARB_R_SPEC:
        eAggHealth := eOutOfSpec;             // 聚合结论：超出规格 / aggregated out of specification
    DL_HARB_R_OK:
        eAggHealth := eOk;                    // 聚合结论：正常 / aggregated OK
ELSE
    eAggHealth := eUnknown;                   // 未选出或全为未知：结论未知（不遮蔽规则见段 10）/ nothing selected means unknown
END_CASE

// 段 10｜Unknown 不遮蔽复核：已知非 OK 存在时结论不得为未知 / segment 10, unknown must not mask a known fault
IF bAnyKnown AND (eAggHealth = eUnknown) AND (nBestRank = DL_HARB_R_NONE) THEN
    eAggHealth := eOutOfSpec;                 // 存在已知态却无等级：按次严重级保守结论文本 / a known state without a rank is treated conservatively
END_IF
IF bAnyUnknown AND bAnyKnown THEN
    eErr := 16#0003_016A;                     // 信息级：存在未知源但未遮蔽已知故障 / info level, unknown sources did not mask the known state
END_IF

// 段 11｜降级判定：有维护/校验类而无故障类即可运行需安排处理 / segment 11, degraded evaluation
bDegraded := bAnyMaintain AND (NOT bAnyFaultLevel); // 降级 = 需处理但不致命 / degraded means action needed but not critical

// 段 12｜首出锁存：复位沿优先于仲裁，且当拍不重新锁存 / segment 12, first-out latching
IF fbTrigReset.Q THEN
    bFirstLatched := FALSE;                   // 复位清锁存 / reset clears the latch
    uFirstInt := DL_HARB_NONE;                // 索引回哨兵 / index back to the sentinel
    uFirstChInt := DL_HARB_CNT_ZERO;          // 通道回 0 / channel back to zero
ELSIF (NOT bFirstLatched) AND (uBestIdx <> DL_HARB_NONE) AND (nBestRank <> DL_HARB_R_OK) THEN
    uFirstInt := uBestIdx;                    // 锁存首个非 OK 源 / latch the first non-OK source
    uFirstChInt := auChannelId[uBestIdx];     // 锁存其对外通道号（索引已由仲裁保证合法）/ latch its channel id, the index is legal by construction
    bFirstLatched := TRUE;                    // 置锁存位 / set the latch
    IF uSameCnt > 1 THEN
        eErr := 16#0003_016A;                 // 信息级：同拍多源同级别，已按来源索引最小仲裁 / info level, ties resolved by the lowest source index
    END_IF
END_IF

// 段 13｜非法枚举汇总置码（故障级，但不中止聚合）/ segment 13, illegal enumeration summary
IF bIllegalEnum THEN
    eErr := 16#0003_0331;                     // 健康枚举非法故障码 / illegal health enumeration fault id
    bError := TRUE;                           // 置故障标志 / raise the error flag
END_IF

// 段 14｜对外镜像 / segment 14, mirror the latched values to the outputs
uFirstIdx := uFirstInt;                       // 首出索引镜像 / first-out index mirror
uFirstChannel := uFirstChInt;                 // 首出通道镜像 / first-out channel mirror
END_FUNCTION_BLOCK

(* ---- FB_DL_DeviceParamWrite.st ---- *)
(*
    FB_DL_DeviceParamWrite —— 设备参数写回事务
    ------------------------------------------------------------------
    分类      : DL_Device / DeviceAccess
    前缀      : FB_DL_
    版本      : 1.0.0
    溯源      : 设备参数「读 → 比 → 判」三段流程的下半段划分（写回 / 复核 / 回滚）；
                只借流程骨架的分类事实，示例页面未声明许可，故按最严口径处置：
                零代码行、零注释引用；白名单机制、事务状态机、回滚策略、错误分级与
                码位 100% 自有；clean-room 重写，未复制任何闭源厂商源码
    平台      : 纯 IEC 61131-3，CODESYS V3.5+ / TwinCAT 3 / InoProShop 通用
    作者      : 道莅代码库 · PLC编程专家（R19）
    ------------------------------------------------------------------
    功能说明  : 备份快照 → 白名单逐项写 → 读回复核 → 不一致即回滚。
                归属裁定（关闭矩阵勘误 M-E3 的悬置项）：参数写回属设备层——写回是设备访问
                能力，工艺层只应下发语义参数，故本件落在 DL_Device 而非 DL_Process。
                核心防御：① 项数越界即拒绝启动事务，不索引数组；
                ② 白名单外项（只读）绝不写，跳过并计数——写只读项在多数设备上会被静默
                   忽略或引发参数区校验失败，后者会让整块参数失效；
                ③ 写超时转回滚；读回偏差超容差同样转回滚（写进去却没保持住 = 参数区有问题）；
                ④ 回滚失败置 033B 并锁存，禁止自动重试——参数区已不可信须人工介入；
                ⑤ bAbort 中止事务但不触发回滚（中止是人为决策，回滚由调用方再发事务决定）。
                规格补正：物理读写不在本件内完成（零厂商库红线），本件经 afActual 输入取
                设备实际值、经 bWriteNow + uActiveIdx 输出驱动上层 IO/驱动层执行写入——
                派单引脚表未含读回通道，实测无法闭环复核，特此补正三个引脚并在收口报告留档。
    错误码    : 16#0003_0170 白名单外项已跳过（uSkipped 非 0）——信息级，正常防御
                16#0003_0171 预留禁用（信息级，不得挪用）
                16#0003_0339 项数越界（不在 1~16）——故障级，事务不启动且不索引数组
                16#0003_033A 写超时 / 读回复核不一致 / 写值非有限——故障级，已转回滚
                16#0003_033B 回滚失败或状态机兜底——故障级，参数区不可信须人工介入（锁存）
    码位总账  : 16#0003_0170 用 / 16#0003_0171 预留 ｜ 16#0003_0339 用 / 16#0003_033A 用 / 16#0003_033B 用
    状态机    : E_DL_ParamWriteState（eIdle / eBackup / eWrite / eVerify / eRollback / eDone / eFault）
                七态，CASE 含 ELSE 兜底，ELSE 回 eFault 并置故障级 033B。
    采样约定  : fbTrigExec / fbTrigAbort / fbTrigReset 与 fbWrite / fbVerify 五个实例在本体首部
                无条件刷新，绝不放入 IF 或 CASE；tWriteTimeout 覆盖整个写入相与回滚相（不做单相
                复位，否则就要在 CASE 内调用实例，违反周期刷新红线），tVerifyTimeout 覆盖复核相；
                bDone 为单周期脉冲，bRollback 保持锁存直到 bReset。
    修订记录  : 2026-11-16 v1.0.0 首次入库（R19）
*)

(*
    枚举 : E_DL_ParamWriteState —— 参数写回事务状态（本文件为全库唯一属主）
*)
TYPE E_DL_ParamWriteState :
(
    eIdle     := 0,                           // 空闲：无事务 / idle, no transaction
    eBackup   := 1,                           // 备份：抓取写前快照 / backup, capture the pre-write snapshot
    eWrite    := 2,                           // 写入：逐项白名单写 / write, item by item with the whitelist
    eVerify   := 3,                           // 复核：读回比对全部已写项 / verify, compare every written item
    eRollback := 4,                           // 回滚：恢复备份快照 / rollback, restore the backup snapshot
    eDone     := 5,                           // 完成：写入并复核通过 / done, written and verified
    eFault    := 6                            // 故障：事务失败或参数区不可信 / fault, the transaction failed or the parameter area is untrustworthy
);
END_TYPE

FUNCTION_BLOCK FB_DL_DeviceParamWrite
VAR_INPUT
    bEnable         : BOOL;                   // 使能，FALSE 中止并撤 bBusy / enable, FALSE aborts and drops the busy flag
    bExecute        : BOOL;                   // 执行，上升沿启动一次写回事务 / execute, rising edge starts one write transaction
    bAbort          : BOOL;                   // 中止，上升沿中止（不触发回滚）/ abort, rising edge aborts without triggering a rollback
    bReset          : BOOL;                   // 复位，上升沿清故障与 bRollback / reset, rising edge clears the faults and the rollback flag
    auIndex         : ARRAY[0..15] OF UINT;   // 参数索引 [索引]，范围 1~65535 / parameter index [index], range 1~65535
    afWriteValue    : ARRAY[0..15] OF REAL;   // 待写值 [用户单位] / value to write [user unit]
    abWritable      : ARRAY[0..15] OF BOOL;   // 白名单：FALSE = 只读项，禁止写 / whitelist, FALSE means read only and forbidden
    afActual        : ARRAY[0..15] OF REAL;   // 设备实际值（由 IO/驱动层每拍提供，规格补正引脚）[用户单位] / device actual values supplied by the IO layer each cycle, a spec correction pin [user unit]
    uCount          : UINT := 0;              // 有效项数 [项]，范围 1~16 / valid item count [item], range 1~16
    fVerifyTol      : REAL := 0.001;          // 读回值容差 [用户单位]，范围 >= 0（0 = 严格相等，不推荐）/ readback tolerance [user unit], >= 0
    tWriteTimeout   : TIME := T#5S;           // 单项写超时 [ms]，范围 100~60000 / per item write timeout [ms], range 100~60000
    tVerifyTimeout  : TIME := T#5S;           // 读回复核超时 [ms]，范围 100~60000 / verification timeout [ms], range 100~60000
END_VAR
VAR_OUTPUT
    bBusy           : BOOL;                   // 事务进行中 / transaction in progress
    bDone           : BOOL;                   // 全部写入并复核通过（单周期脉冲）/ everything written and verified, a single-cycle pulse
    bRollback       : BOOL;                   // 发生过回滚（锁存）/ a rollback occurred, latched
    uWritten        : UINT;                   // 实际写入并复核通过的项数 [项] / items written and verified [item]
    uSkipped        : UINT;                   // 因白名单或非法索引被跳过的项数 [项] / items skipped due to the whitelist or an illegal index [item]
    uFailedIdx      : UINT;                   // 首个失败项索引，16#FFFF = 无 [索引] / first failed item index, sentinel 16#FFFF when none [index]
    afReadback      : ARRAY[0..15] OF REAL;   // 复核读回值 [用户单位] / verification readback values [user unit]
    uActiveIdx      : UINT;                   // 当前事务活动项索引（供 IO 层定位，规格补正引脚）[索引] / active item index for the IO layer, a spec correction pin [index]
    bWriteNow       : BOOL;                   // 本拍请求 IO 层执行写入/回写（规格补正引脚）/ request the IO layer to perform the write or the restore in this cycle, a spec correction pin
    eErr            : UDINT;                  // 错误码，0=正常 / error id, 0=ok
    bError          : BOOL;                   // 故障标志，eErr 为故障级时 TRUE / error flag, TRUE on fault-level eErr
END_VAR
VAR
    eState          : E_DL_ParamWriteState := eIdle; // 状态机当前态 / current state machine state
    fbTrigExec      : R_TRIG;                 // 执行沿实例，本体首部无条件刷新 / execute edge instance, refreshed unconditionally
    fbTrigAbort     : R_TRIG;                 // 中止沿实例，本体首部无条件刷新 / abort edge instance, refreshed unconditionally
    fbTrigReset     : R_TRIG;                 // 复位沿实例，本体首部无条件刷新 / reset edge instance, refreshed unconditionally
    fbWrite         : TON;                    // 写超时实例，本体首部无条件刷新 / write timeout instance, refreshed unconditionally
    fbVerify        : TON;                    // 复核超时实例，本体首部无条件刷新 / verification timeout instance, refreshed unconditionally
    uIdx            : UINT;                   // 事务游标 [索引]，范围 0~15 / transaction cursor [index], range 0~15
    uScan           : UINT;                   // 全表扫描游标 [索引] / full table scan cursor [index]
    afBackup        : ARRAY[0..15] OF REAL;   // 写前快照 [用户单位] / pre-write snapshot [user unit]
    bAllOk         : BOOL;                    // 全表一致性判定标志 / full table consistency flag
    bItemOk        : BOOL;                    // 单项一致性判定标志 / single item consistency flag
    bNonFin        : BOOL;                    // 写值非有限判定标志 / non-finite write value flag
    fTolEff        : REAL;                    // 生效容差（负值收敛到 0）[用户单位] / effective tolerance, negatives converge to zero [user unit]
END_VAR
VAR CONSTANT
    DL_DPW_ITEM_MAX  : UINT := 16;            // 项数上限 [项] / item count upper bound [item]
    DL_DPW_NONE      : UINT := 16#FFFF;       // 无失败项哨兵 [索引] / no failed item sentinel [index]
    DL_DPW_TMO_MIN   : TIME := T#100MS;       // 超时下限 [ms] / timeout lower bound [ms]
    DL_DPW_TMO_MAX   : TIME := T#60S;         // 超时上限 [ms] / timeout upper bound [ms]
    DL_DPW_CNT_MAX   : UINT := 65535;         // 项数计数饱和值 [项] / item counter saturation value [item]
    DL_FLOAT_EPS     : REAL := 1.0E-6;        // 浮点判等容差 [无量纲] / float equality tolerance [dimensionless]
    DL_DPW_INF_GUARD : REAL := 1.0E38;        // 非有限幅值判定阈值 [无量纲] / non-finite magnitude guard [dimensionless]
    DL_DPW_ZERO      : REAL := 0.0;           // 零值常量，避免裸字面量 [无量纲] / zero constant, avoids a bare literal [dimensionless]
    DL_DPW_CNT_ZERO  : UINT := 0;             // 无符号零常量 [无量纲] / unsigned zero constant [dimensionless]
END_VAR

// 段 1｜边沿与定时器实例无条件周期刷新（红线：严禁放入条件分支）/ segment 1, unconditional refresh
fbTrigExec(CLK := bExecute);
fbTrigAbort(CLK := bAbort);
fbTrigReset(CLK := bReset);
fbWrite(IN := (eState = eWrite) OR (eState = eRollback), PT := tWriteTimeout); // 写入与回写共用写超时 / writing and restoring share the write timeout
fbVerify(IN := (eState = eVerify), PT := tVerifyTimeout);                      // 复核独立超时 / verification has its own timeout

// 段 2｜输出与错误状态预置（bRollback 为保持量，不预置）/ segment 2, preset outputs, the rollback latch is kept
bDone := FALSE;                               // 单周期脉冲先清 / clear the single-cycle pulse first
bWriteNow := FALSE;                           // 写请求先清 / clear the write request
eErr := 0;                                    // 预置无错误 / preset no error
bError := FALSE;                              // 预置无故障 / preset no fault
bBusy := (eState <> eIdle) AND (eState <> eDone) AND (eState <> eFault); // 忙标志由状态导出 / the busy flag derives from the state

// 段 3｜复位沿清故障与回滚锁存 / segment 3, reset clears the faults and the rollback latch
IF fbTrigReset.Q THEN
    bRollback := FALSE;                       // 清回滚锁存 / clear the rollback latch
    uFailedIdx := DL_DPW_NONE;                // 清失败项索引 / clear the failed item index
    IF (eState = eFault) OR (eState = eDone) THEN
        eState := eIdle;                      // 复位允许离开故障与完成态 / a reset leaves the fault and done states
    END_IF
END_IF

// 段 4｜中止沿：人为中止不置故障、不自动回滚 / segment 4, abort without a fault and without a rollback
IF fbTrigAbort.Q THEN
    eState := eIdle;                          // 回空闲态 / back to idle
    bBusy := FALSE;                           // 撤忙标志 / drop the busy flag
    bWriteNow := FALSE;                       // 撤写请求 / drop the write request
    RETURN;                                   // 中止即出口 / abort is the exit
END_IF

// 段 5｜使能闸 / segment 5, enable gate
IF NOT bEnable THEN
    eState := eIdle;                          // 回空闲态 / back to idle
    bBusy := FALSE;                           // 撤忙标志 / drop the busy flag
    RETURN;                                   // 失能即出口 / disabled is the exit
END_IF

// 段 6｜容差收敛与参数闸（超时与容差先口径统一）/ segment 6, tolerance and timeout convergence
fTolEff := MAX(fVerifyTol, DL_DPW_ZERO);      // 容差负数收敛到 0（0 = 严格相等，不推荐）/ a negative tolerance converges to zero
IF (tWriteTimeout < DL_DPW_TMO_MIN) OR (tWriteTimeout > DL_DPW_TMO_MAX)
   OR (tVerifyTimeout < DL_DPW_TMO_MIN) OR (tVerifyTimeout > DL_DPW_TMO_MAX) THEN
    eErr := 16#0003_0339;                     // 超时参数越界按项数同码处理（事务不可启动）/ an illegal timeout shares the item count fault id, the transaction cannot start
    bError := TRUE;                           // 置故障标志 / raise the error flag
    eState := eFault;                         // 落故障态 / enter the fault state
    bBusy := FALSE;                           // 不忙 / not busy
    RETURN;                                   // 故障级提前返回 / early return on fault
END_IF

// 段 7｜执行沿启动：项数闸在最前，越界绝不索引数组 / segment 7, start edge with the item count gate first
IF fbTrigExec.Q AND ((eState = eIdle) OR (eState = eDone) OR (eState = eFault)) THEN
    IF (uCount < 1) OR (uCount > DL_DPW_ITEM_MAX) THEN
        eErr := 16#0003_0339;                 // 项数越界故障码 / item count out of range fault id
        bError := TRUE;                       // 置故障标志 / raise the error flag
        eState := eFault;                     // 落故障态 / enter the fault state
        RETURN;                               // 事务不启动 / the transaction never starts
    END_IF
    uIdx := DL_DPW_CNT_ZERO;                  // 游标归零 / reset the cursor
    uWritten := DL_DPW_CNT_ZERO;              // 已写项数清零 / clear the written count
    uSkipped := DL_DPW_CNT_ZERO;              // 跳过项数清零 / clear the skipped count
    uFailedIdx := DL_DPW_NONE;                // 失败项清哨兵 / reset the failed item to the sentinel
    uActiveIdx := DL_DPW_NONE;                // 活动项清哨兵 / reset the active index to the sentinel
    eState := eBackup;                        // 进入备份相 / enter the backup phase
END_IF

// 段 8｜状态机（含 ELSE 兜底）/ segment 8, state machine with ELSE fallback
CASE eState OF
    eIdle:
        bBusy := FALSE;                       // 空闲不忙 / idle is not busy

    eBackup:
        // 段 9｜抓取写前快照（白名单外项也备份，回滚需要完整镜像）/ segment 9, capture the pre-write snapshot
        FOR uScan := 0 TO uCount - 1 DO
            afBackup[uScan] := afActual[uScan]; // 快照取设备实际值 / the snapshot takes the device actual value
            afReadback[uScan] := afActual[uScan]; // 读回镜像同步初始化 / initialise the readback mirror
        END_FOR
        eState := eWrite;                     // 备份完成进入写入相 / the backup is complete, enter the write phase

    eWrite:
        // 段 10｜逐项白名单写：只读项绝不写，跳过并计数 / segment 10, whitelisted writes only
        IF uIdx >= uCount THEN
            eState := eVerify;                // 全部处理完进入复核相 / everything processed, enter the verification phase
        ELSE
            bNonFin := (afWriteValue[uIdx] <> afWriteValue[uIdx])
                    OR (afWriteValue[uIdx] > DL_DPW_INF_GUARD)
                    OR (afWriteValue[uIdx] < -DL_DPW_INF_GUARD); // 写值非有限判定 / non-finite write value detection
            IF bNonFin THEN
                eErr := 16#0003_033A;         // 写值非有限，转回滚 / a non-finite value triggers the rollback
                bError := TRUE;               // 置故障标志 / raise the error flag
                uFailedIdx := uIdx;           // 记录失败项 / record the failed item
                eState := eRollback;          // 转回滚相 / enter the rollback phase
            ELSIF (NOT abWritable[uIdx]) OR (auIndex[uIdx] < 1) THEN
                IF uSkipped < DL_DPW_CNT_MAX THEN
                    uSkipped := uSkipped + 1; // 白名单外或索引非法：饱和计数跳过 / outside the whitelist or an illegal index, saturating skip count
                END_IF
                eErr := 16#0003_0170;         // 信息级：白名单外项已跳过 / info level, the item was skipped
                uIdx := uIdx + 1;             // 游标前进 / advance the cursor
            ELSE
                uActiveIdx := uIdx;           // 发布活动项 / publish the active item
                bWriteNow := TRUE;            // 请求 IO 层执行写入 / request the IO layer to write
                afReadback[uIdx] := afActual[uIdx]; // 同步读回镜像 / keep the readback mirror in step
                bItemOk := ABS(afActual[uIdx] - afWriteValue[uIdx]) <= fTolEff; // 单项落值判定 / single item settled test
                IF bItemOk THEN
                    uWritten := uWritten + 1; // 落值即计入已写 / a settled value counts as written
                    uIdx := uIdx + 1;         // 游标前进（超时按整个写入相计，避免在 CASE 内调用实例）/ advance the cursor, the timeout covers the whole write phase so no instance call lives inside CASE
                ELSIF fbWrite.Q THEN
                    eErr := 16#0003_033A;     // 写超时，转回滚 / a write timeout triggers the rollback
                    bError := TRUE;           // 置故障标志 / raise the error flag
                    uFailedIdx := uIdx;       // 记录失败项 / record the failed item
                    eState := eRollback;      // 转回滚相 / enter the rollback phase
                END_IF
            END_IF
        END_IF

    eVerify:
        // 段 11｜全表复核：读回值与目标值逐项比对（只读项不参与）/ segment 11, full table verification
        bAllOk := TRUE;                       // 先假设一致 / assume consistency first
        FOR uScan := 0 TO uCount - 1 DO
            IF abWritable[uScan] AND (auIndex[uScan] >= 1) THEN
                afReadback[uScan] := afActual[uScan]; // 抓取复核读回值 / capture the verification readback
                IF ABS(afActual[uScan] - afWriteValue[uScan]) > fTolEff THEN
                    bAllOk := FALSE;          // 任一项不一致即失败 / a single mismatch fails the verification
                    uFailedIdx := uScan;      // 记录首个不一致项 / record the first mismatching item
                END_IF
            END_IF
        END_FOR
        IF bAllOk THEN
            eState := eDone;                  // 复核通过 / verification passed
            bDone := TRUE;                    // 单周期完成脉冲 / single-cycle done pulse
            bBusy := FALSE;                   // 事务结束 / the transaction finished
        ELSIF fbVerify.Q THEN
            eErr := 16#0003_033A;             // 复核不一致且超时，转回滚 / verification failed within its timeout, roll back
            bError := TRUE;                   // 置故障标志 / raise the error flag
            eState := eRollback;              // 转回滚相 / enter the rollback phase
        ELSE
            bBusy := TRUE;                    // 复核进行中 / verification in progress
        END_IF

    eRollback:
        // 段 12｜回滚：把备份快照逐项写回，全表恢复才算出清 / segment 12, restore the snapshot
        bAllOk := TRUE;                       // 先假设已恢复 / assume restored first
        bWriteNow := TRUE;                    // 持续请求 IO 层回写 / keep requesting the restore
        FOR uScan := 0 TO uCount - 1 DO
            IF abWritable[uScan] AND (auIndex[uScan] >= 1) THEN
                uActiveIdx := uScan;          // 回写活动项 / the item being restored
                IF ABS(afActual[uScan] - afBackup[uScan]) > fTolEff THEN
                    bAllOk := FALSE;          // 尚未恢复 / not yet restored
                    uFailedIdx := uScan;      // 记录回滚受阻项 / record the blocked item
                END_IF
                afReadback[uScan] := afActual[uScan]; // 同步读回 / keep the readback in step
            END_IF
        END_FOR
        IF bAllOk THEN
            bRollback := TRUE;                // 回滚完成，锁存 / the rollback completed, latch it
            eErr := 16#0003_033A;             // 事务失败（已回滚）故障码 / the transaction failed and was rolled back
            bError := TRUE;                   // 置故障标志 / raise the error flag
            eState := eFault;                 // 进故障态待人工确认 / enter the fault state pending manual acknowledgement
            bWriteNow := FALSE;               // 撤回写请求 / drop the restore request
        ELSIF fbWrite.Q THEN
            bRollback := TRUE;                // 回滚失败同样锁存 / a failed rollback is latched as well
            eErr := 16#0003_033B;             // 参数区不可信，禁止自动重试 / the parameter area is untrustworthy, no automatic retry
            bError := TRUE;                   // 置故障标志 / raise the error flag
            eState := eFault;                 // 进故障态锁存 / latch the fault state
            bWriteNow := FALSE;               // 撤回写请求 / drop the restore request
        END_IF

    eDone:
        bBusy := FALSE;                       // 完成态不忙 / the done state is not busy
        bWriteNow := FALSE;                   // 撤写请求 / drop the write request

    eFault:
        bBusy := FALSE;                       // 故障态不忙 / the fault state is not busy
        bWriteNow := FALSE;                   // 撤写请求 / drop the write request

ELSE
    eErr := 16#0003_033B;                     // 故障级：非法状态兜底 / fault level, illegal state fallback
    bError := TRUE;                           // 置故障标志 / raise the error flag
    eState := eFault;                         // 回故障态 / fall back to the fault state
    bWriteNow := FALSE;                       // 撤写请求，绝不留在写入状态 / drop the write request, never stay in a writing state
END_CASE
END_FUNCTION_BLOCK
